//     Drive/Inputs/In/nState1 @bit 4 <-> STM Status/Status/Moving positive
//     Drive/Inputs/In/nState1 @bit 1 <-> STM Status/Status/Ready
//     Drive/Inputs/In/nState1 <-> STM Status/Status/Ready to enable
//     Drive/Inputs/In/nState1 @bit 6 <-> STM Status/Status/Torque reduced
//     Drive/Inputs/In/nState1 @bit 2 <-> STM Status/Status/Warning
//     Drive/Inputs/In/nState2 @bit 3 <-> STM Status/Status/Digital input 1
//     Drive/Inputs/In/nState2 @bit 4 <-> STM Status/Status/Digital input 2
//     Drive/Inputs/In/nState2 @bit 5 <-> STM Status/Status/Sync error
//     Drive/Inputs/In/nState2 @bit 7 <-> STM Status/Status/TxPDO Toggle
//     Drive/Inputs/In/nState4 @bit 1 <-> WcState/InputToggle
//     Drive/Inputs/In/nState4 <-> WcState/WcState
//     Drive/Outputs/Out/nCtrl1 <-> STM Control/Control/Enable
//     Drive/Outputs/Out/nCtrl1 @bit 2 <-> STM Control/Control/Reduce torque
//     Drive/Outputs/Out/nCtrl1 @bit 1 <-> STM Control/Control/Reset
//     Drive/Outputs/Out/nDataOut2[0] <-> STM Velocity/Velocity
//   (this object) <-> PLC Rail (EtherCAT)/Power (EK1200)/PLC Junction 2 (EK1122)/X1 HXR EC1 (EK1100)/EC1 E2 (EK1122)/X1 IM2L0-XTES (EK1100)/IM2L0-EL5042
//     Enc/Inputs/In/nComState @bit 1 <-> WcState/InputToggle
//     Enc/Inputs/In/nComState <-> WcState/WcState
//     Enc/Inputs/In/nDataIn1 <-> FB Inputs Channel 1/Position
//     Enc/Inputs/In/nState1 @bit 12 <-> FB Inputs Channel 1/Status/Diag
//     Enc/Inputs/In/nState1 @bit 1 <-> FB Inputs Channel 1/Status/Error
//     Enc/Inputs/In/nState1 @bit 14 <-> FB Inputs Channel 1/Status/Input cycle counter
//     Enc/Inputs/In/nState1 @bit 2 <-> FB Inputs Channel 1/Status/Ready
//     Enc/Inputs/In/nState1 @bit 13 <-> FB Inputs Channel 1/Status/TxPDO State
//     Enc/Inputs/In/nState1 <-> FB Inputs Channel 1/Status/Warning
//   (this object) <-> PLC Rail (EtherCAT)/Power (EK1200)/PLC Junction 2 (EK1122)/X1 HXR EC1 (EK1100)/EC1 E2 (EK1122)/X1 IM2L0-XTES (EK1100)/IM2L0-EL7041
//     Drive/Inputs/In/nState1 @bit 3 <-> STM Status/Status/Error
//     Drive/Inputs/In/nState1 @bit 5 <-> STM Status/Status/Moving negative
//     Drive/Inputs/In/nState1 @bit 4 <-> STM Status/Status/Moving positive
//     Drive/Inputs/In/nState1 @bit 1 <-> STM Status/Status/Ready
//     Drive/Inputs/In/nState1 <-> STM Status/Status/Ready to enable
//     Drive/Inputs/In/nState1 @bit 6 <-> STM Status/Status/Torque reduced
//     Drive/Inputs/In/nState1 @bit 2 <-> STM Status/Status/Warning
//     Drive/Inputs/In/nState2 @bit 3 <-> STM Status/Status/Digital input 1
//     Drive/Inputs/In/nState2 @bit 4 <-> STM Status/Status/Digital input 2
//     Drive/Inputs/In/nState2 @bit 5 <-> STM Status/Status/Sync error
//     Drive/Inputs/In/nState2 @bit 7 <-> STM Status/Status/TxPDO Toggle
//     Drive/Inputs/In/nState4 @bit 1 <-> WcState/InputToggle
//     Drive/Inputs/In/nState4 <-> WcState/WcState
//     Drive/Outputs/Out/nCtrl1 <-> STM Control/Control/Enable
//     Drive/Outputs/Out/nCtrl1 @bit 2 <-> STM Control/Control/Reduce torque
//     Drive/Outputs/Out/nCtrl1 @bit 1 <-> STM Control/Control/Reset
//     Drive/Outputs/Out/nDataOut2[0] <-> STM Velocity/Velocity
//   (this object) <-> PLC Rail (EtherCAT)/Power (EK1200)/PLC Junction 2 (EK1122)/X1 HXR EC1 (EK1100)/EC1 E2 (EK1122)/X1 IM2L0-XTES (EK1100)/IM2L0-EL7342
//     Drive/Inputs/In/nState1 @bit 3 <-> DCM Status Channel 1/Status/Error
//     Drive/Inputs/In/nState1 @bit 3 <-> DCM Status Channel 2/Status/Error
//     Drive/Inputs/In/nState1 @bit 5 <-> DCM Status Channel 1/Status/Moving negative
//     Drive/Inputs/In/nState1 @bit 5 <-> DCM Status Channel 2/Status/Moving negative
//     Drive/Inputs/In/nState1 @bit 4 <-> DCM Status Channel 1/Status/Moving positive
//     Drive/Inputs/In/nState1 @bit 4 <-> DCM Status Channel 2/Status/Moving positive
//     Drive/Inputs/In/nState1 @bit 1 <-> DCM Status Channel 1/Status/Ready
//     Drive/Inputs/In/nState1 @bit 1 <-> DCM Status Channel 2/Status/Ready
//     Drive/Inputs/In/nState1 <-> DCM Status Channel 1/Status/Ready to enable
//     Drive/Inputs/In/nState1 <-> DCM Status Channel 2/Status/Ready to enable
//     Drive/Inputs/In/nState1 @bit 6 <-> DCM Status Channel 1/Status/Torque reduced
//     Drive/Inputs/In/nState1 @bit 6 <-> DCM Status Channel 2/Status/Torque reduced
//     Drive/Inputs/In/nState1 @bit 2 <-> DCM Status Channel 1/Status/Warning
//     Drive/Inputs/In/nState1 @bit 2 <-> DCM Status Channel 2/Status/Warning
//     Drive/Inputs/In/nState2 @bit 3 <-> DCM Status Channel 1/Status/Digital input 1
//     Drive/Inputs/In/nState2 @bit 4 <-> DCM Status Channel 1/Status/Digital input 2
//     Drive/Inputs/In/nState2 @bit 3 <-> DCM Status Channel 2/Status/Digital input 1
//     Drive/Inputs/In/nState2 @bit 4 <-> DCM Status Channel 2/Status/Digital input 2
//     Drive/Inputs/In/nState2 @bit 5 <-> DCM Status Channel 1/Status/Sync error
//     Drive/Inputs/In/nState2 @bit 5 <-> DCM Status Channel 2/Status/Sync error
//     Drive/Inputs/In/nState2 @bit 7 <-> DCM Status Channel 1/Status/TxPDO Toggle
//     Drive/Inputs/In/nState2 @bit 7 <-> DCM Status Channel 2/Status/TxPDO Toggle
//     Drive/Inputs/In/nState4 @bit 1 <-> WcState/InputToggle
//     Drive/Inputs/In/nState4 <-> WcState/WcState
//     Drive/Outputs/Out/nCtrl1 <-> DCM Control Channel 1/Control/Enable
//     Drive/Outputs/Out/nCtrl1 <-> DCM Control Channel 2/Control/Enable
//     Drive/Outputs/Out/nCtrl1 @bit 2 <-> DCM Control Channel 1/Control/Reduce torque
//     Drive/Outputs/Out/nCtrl1 @bit 2 <-> DCM Control Channel 2/Control/Reduce torque
//     Drive/Outputs/Out/nCtrl1 @bit 1 <-> DCM Control Channel 1/Control/Reset
//     Drive/Outputs/Out/nCtrl1 @bit 1 <-> DCM Control Channel 2/Control/Reset
//     Drive/Outputs/Out/nCtrl1 @bit 3 <-> DCM Control Channel 1/Control/Threshold active
//     Drive/Outputs/Out/nCtrl1 @bit 3 <-> DCM Control Channel 2/Control/Threshold active
//     Drive/Outputs/Out/nDataOut2[0] <-> DCM Velocity Channel 1/Velocity
//     Drive/Outputs/Out/nDataOut2[0] <-> DCM Velocity Channel 2/Velocity
//     Enc/Inputs/In/nDataIn1[0] <-> ENC Status compact Channel 1/Counter value
//     Enc/Inputs/In/nDataIn1[0] <-> ENC Status compact Channel 2/Counter value
//     Enc/Inputs/In/nDataIn2[0] <-> ENC Status compact Channel 1/Latch value
//     Enc/Inputs/In/nDataIn2[0] <-> ENC Status compact Channel 2/Latch value
//     Enc/Inputs/In/nState1 @bit 4 <-> ENC Status compact Channel 1/Status/Counter overflow
//     Enc/Inputs/In/nState1 @bit 4 <-> ENC Status compact Channel 2/Status/Counter overflow
//     Enc/Inputs/In/nState1 @bit 3 <-> ENC Status compact Channel 1/Status/Counter underflow
//     Enc/Inputs/In/nState1 @bit 3 <-> ENC Status compact Channel 2/Status/Counter underflow
//     Enc/Inputs/In/nState1 @bit 7 <-> ENC Status compact Channel 1/Status/Extrapolation stall
//     Enc/Inputs/In/nState1 @bit 7 <-> ENC Status compact Channel 2/Status/Extrapolation stall
//     Enc/Inputs/In/nState1 @bit 1 <-> ENC Status compact Channel 1/Status/Latch extern valid
//     Enc/Inputs/In/nState1 @bit 1 <-> ENC Status compact Channel 2/Status/Latch extern valid
//     Enc/Inputs/In/nState1 @bit 2 <-> ENC Status compact Channel 1/Status/Set counter done
//     Enc/Inputs/In/nState1 @bit 2 <-> ENC Status compact Channel 2/Status/Set counter done
//     Enc/Inputs/In/nState2 @bit 4 <-> ENC Status compact Channel 1/Status/Status of extern latch
//     Enc/Inputs/In/nState2 @bit 4 <-> ENC Status compact Channel 2/Status/Status of extern latch
//     Enc/Inputs/In/nState2 <-> ENC Status compact Channel 1/Status/Status of input A
//     Enc/Inputs/In/nState2 <-> ENC Status compact Channel 2/Status/Status of input A
//     Enc/Inputs/In/nState2 @bit 1 <-> ENC Status compact Channel 1/Status/Status of input B
//     Enc/Inputs/In/nState2 @bit 1 <-> ENC Status compact Channel 2/Status/Status of input B
//     Enc/Inputs/In/nState2 @bit 5 <-> ENC Status compact Channel 1/Status/Sync error
//     Enc/Inputs/In/nState2 @bit 5 <-> ENC Status compact Channel 2/Status/Sync error
//     Enc/Inputs/In/nState2 @bit 7 <-> ENC Status compact Channel 1/Status/TxPDO Toggle
//     Enc/Inputs/In/nState2 @bit 7 <-> ENC Status compact Channel 2/Status/TxPDO Toggle
//     Enc/Inputs/In/nState4 @bit 1 <-> WcState/InputToggle
//     Enc/Inputs/In/nState4 <-> WcState/WcState
//     Enc/Outputs/Out/nCtrl1 @bit 3 <-> ENC Control compact Channel 1/Control/Enable latch extern on negative edge
//     Enc/Outputs/Out/nCtrl1 @bit 3 <-> ENC Control compact Channel 2/Control/Enable latch extern on negative edge
//     Enc/Outputs/Out/nCtrl1 @bit 1 <-> ENC Control compact Channel 1/Control/Enable latch extern on positive edge
//     Enc/Outputs/Out/nCtrl1 @bit 1 <-> ENC Control compact Channel 2/Control/Enable latch extern on positive edge
//     Enc/Outputs/Out/nCtrl1 @bit 2 <-> ENC Control compact Channel 1/Control/Set counter
//     Enc/Outputs/Out/nCtrl1 @bit 2 <-> ENC Control compact Channel 2/Control/Set counter
//     Enc/Outputs/Out/nDataOut1[0] <-> ENC Control compact Channel 1/Set counter value
//     Enc/Outputs/Out/nDataOut1[0] <-> ENC Control compact Channel 2/Set counter value
//   (this object) <-> PLC Rail (EtherCAT)/Power (EK1200)/PLC Junction 2 (EK1122)/X2 HXR EC2 (EK1100)/EC2 E1 (EK1122)/X1 IM3L0-PPM (EK1100)/IM3L0-EL5042
//     Enc/Inputs/In/nComState @bit 1 <-> WcState/InputToggle
//     Enc/Inputs/In/nComState <-> WcState/WcState
//     Enc/Inputs/In/nDataIn1 <-> FB Inputs Channel 1/Position
//     Enc/Inputs/In/nState1 @bit 12 <-> FB Inputs Channel 1/Status/Diag
//     Enc/Inputs/In/nState1 @bit 1 <-> FB Inputs Channel 1/Status/Error
//     Enc/Inputs/In/nState1 @bit 14 <-> FB Inputs Channel 1/Status/Input cycle counter
//     Enc/Inputs/In/nState1 @bit 2 <-> FB Inputs Channel 1/Status/Ready
//     Enc/Inputs/In/nState1 @bit 13 <-> FB Inputs Channel 1/Status/TxPDO State
//     Enc/Inputs/In/nState1 <-> FB Inputs Channel 1/Status/Warning
//   (this object) <-> PLC Rail (EtherCAT)/Power (EK1200)/PLC Junction 2 (EK1122)/X2 HXR EC2 (EK1100)/EC2 E1 (EK1122)/X1 IM3L0-PPM (EK1100)/IM3L0-EL7041
//     Drive/Inputs/In/nState1 @bit 3 <-> STM Status/Status/Error
//     Drive/Inputs/In/nState1 @bit 5 <-> STM Status/Status/Moving negative
//     Drive/Inputs/In/nState1 @bit 4 <-> STM Status/Status/Moving positive
//     Drive/Inputs/In/nState1 @bit 1 <-> STM Status/Status/Ready
//     Drive/Inputs/In/nState1 <-> STM Status/Status/Ready to enable
//     Drive/Inputs/In/nState1 @bit 6 <-> STM Status/Status/Torque reduced
//     Drive/Inputs/In/nState1 @bit 2 <-> STM Status/Status/Warning
//     Drive/Inputs/In/nState2 @bit 3 <-> STM Status/Status/Digital input 1
//     Drive/Inputs/In/nState2 @bit 4 <-> STM Status/Status/Digital input 2
//     Drive/Inputs/In/nState2 @bit 5 <-> STM Status/Status/Sync error
//     Drive/Inputs/In/nState2 @bit 7 <-> STM Status/Status/TxPDO Toggle
//     Drive/Inputs/In/nState4 @bit 1 <-> WcState/InputToggle
//     Drive/Inputs/In/nState4 <-> WcState/WcState
//     Drive/Outputs/Out/nCtrl1 <-> STM Control/Control/Enable
//     Drive/Outputs/Out/nCtrl1 @bit 2 <-> STM Control/Control/Reduce torque
//     Drive/Outputs/Out/nCtrl1 @bit 1 <-> STM Control/Control/Reset
//     Drive/Outputs/Out/nDataOut2[0] <-> STM Velocity/Velocity
//   (this object) <-> PLC Rail (EtherCAT)/Power (EK1200)/PLC Junction 2 (EK1122)/X2 HXR EC2 (EK1100)/EC2 E2 (EK1122)/X1 IM4L0-XTES (EK1100)/IM4L0-EL5042
//     Enc/Inputs/In/nComState @bit 1 <-> WcState/InputToggle
//     Enc/Inputs/In/nComState <-> WcState/WcState
//     Enc/Inputs/In/nDataIn1 <-> FB Inputs Channel 1/Position
//     Enc/Inputs/In/nState1 @bit 12 <-> FB Inputs Channel 1/Status/Diag
//     Enc/Inputs/In/nState1 @bit 1 <-> FB Inputs Channel 1/Status/Error
//     Enc/Inputs/In/nState1 @bit 14 <-> FB Inputs Channel 1/Status/Input cycle counter
//     Enc/Inputs/In/nState1 @bit 2 <-> FB Inputs Channel 1/Status/Ready
//     Enc/Inputs/In/nState1 @bit 13 <-> FB Inputs Channel 1/Status/TxPDO State
//     Enc/Inputs/In/nState1 <-> FB Inputs Channel 1/Status/Warning
//   (this object) <-> PLC Rail (EtherCAT)/Power (EK1200)/PLC Junction 2 (EK1122)/X2 HXR EC2 (EK1100)/EC2 E2 (EK1122)/X1 IM4L0-XTES (EK1100)/IM4L0-EL7041
//     Drive/Inputs/In/nState1 @bit 3 <-> STM Status/Status/Error
//     Drive/Inputs/In/nState1 @bit 5 <-> STM Status/Status/Moving negative
//     Drive/Inputs/In/nState1 @bit 4 <-> STM Status/Status/Moving positive
//     Drive/Inputs/In/nState1 @bit 1 <-> STM Status/Status/Ready
//     Drive/Inputs/In/nState1 <-> STM Status/Status/Ready to enable
//     Drive/Inputs/In/nState1 @bit 6 <-> STM Status/Status/Torque reduced
//     Drive/Inputs/In/nState1 @bit 2 <-> STM Status/Status/Warning
//     Drive/Inputs/In/nState2 @bit 3 <-> STM Status/Status/Digital input 1
//     Drive/Inputs/In/nState2 @bit 4 <-> STM Status/Status/Digital input 2
//     Drive/Inputs/In/nState2 @bit 5 <-> STM Status/Status/Sync error
//     Drive/Inputs/In/nState2 @bit 7 <-> STM Status/Status/TxPDO Toggle
//     Drive/Inputs/In/nState4 @bit 1 <-> WcState/InputToggle
//     Drive/Inputs/In/nState4 <-> WcState/WcState
//     Drive/Outputs/Out/nCtrl1 <-> STM Control/Control/Enable
//     Drive/Outputs/Out/nCtrl1 @bit 2 <-> STM Control/Control/Reduce torque
//     Drive/Outputs/Out/nCtrl1 @bit 1 <-> STM Control/Control/Reset
//     Drive/Outputs/Out/nDataOut2[0] <-> STM Velocity/Velocity
//   (this object) <-> PLC Rail (EtherCAT)/Power (EK1200)/PLC Junction 2 (EK1122)/X2 HXR EC2 (EK1100)/EC2 E2 (EK1122)/X1 IM4L0-XTES (EK1100)/IM4L0-EL7342
//     Drive/Inputs/In/nState1 @bit 3 <-> DCM Status Channel 1/Status/Error
//     Drive/Inputs/In/nState1 @bit 3 <-> DCM Status Channel 2/Status/Error
//     Drive/Inputs/In/nState1 @bit 5 <-> DCM Status Channel 1/Status/Moving negative
//     Drive/Inputs/In/nState1 @bit 5 <-> DCM Status Channel 2/Status/Moving negative
//     Drive/Inputs/In/nState1 @bit 4 <-> DCM Status Channel 1/Status/Moving positive
//     Drive/Inputs/In/nState1 @bit 4 <-> DCM Status Channel 2/Status/Moving positive
//     Drive/Inputs/In/nState1 @bit 1 <-> DCM Status Channel 1/Status/Ready
//     Drive/Inputs/In/nState1 @bit 1 <-> DCM Status Channel 2/Status/Ready
//     Drive/Inputs/In/nState1 <-> DCM Status Channel 1/Status/Ready to enable
//     Drive/Inputs/In/nState1 <-> DCM Status Channel 2/Status/Ready to enable
//     Drive/Inputs/In/nState1 @bit 6 <-> DCM Status Channel 1/Status/Torque reduced
//     Drive/Inputs/In/nState1 @bit 6 <-> DCM Status Channel 2/Status/Torque reduced
//     Drive/Inputs/In/nState1 @bit 2 <-> DCM Status Channel 1/Status/Warning
//     Drive/Inputs/In/nState1 @bit 2 <-> DCM Status Channel 2/Status/Warning
//     Drive/Inputs/In/nState2 @bit 3 <-> DCM Status Channel 1/Status/Digital input 1
//     Drive/Inputs/In/nState2 @bit 4 <-> DCM Status Channel 1/Status/Digital input 2
//     Drive/Inputs/In/nState2 @bit 3 <-> DCM Status Channel 2/Status/Digital input 1
//     Drive/Inputs/In/nState2 @bit 4 <-> DCM Status Channel 2/Status/Digital input 2
//     Drive/Inputs/In/nState2 @bit 5 <-> DCM Status Channel 1/Status/Sync error
//     Drive/Inputs/In/nState2 @bit 5 <-> DCM Status Channel 2/Status/Sync error
//     Drive/Inputs/In/nState2 @bit 7 <-> DCM Status Channel 1/Status/TxPDO Toggle
//     Drive/Inputs/In/nState2 @bit 7 <-> DCM Status Channel 2/Status/TxPDO Toggle
//     Drive/Inputs/In/nState4 @bit 1 <-> WcState/InputToggle
//     Drive/Inputs/In/nState4 <-> WcState/WcState
//     Drive/Outputs/Out/nCtrl1 <-> DCM Control Channel 1/Control/Enable
//     Drive/Outputs/Out/nCtrl1 <-> DCM Control Channel 2/Control/Enable
//     Drive/Outputs/Out/nCtrl1 @bit 2 <-> DCM Control Channel 1/Control/Reduce torque
//     Drive/Outputs/Out/nCtrl1 @bit 2 <-> DCM Control Channel 2/Control/Reduce torque
//     Drive/Outputs/Out/nCtrl1 @bit 1 <-> DCM Control Channel 1/Control/Reset
//     Drive/Outputs/Out/nCtrl1 @bit 1 <-> DCM Control Channel 2/Control/Reset
//     Drive/Outputs/Out/nCtrl1 @bit 3 <-> DCM Control Channel 1/Control/Threshold active
//     Drive/Outputs/Out/nCtrl1 @bit 3 <-> DCM Control Channel 2/Control/Threshold active
//     Drive/Outputs/Out/nDataOut2[0] <-> DCM Velocity Channel 1/Velocity
//     Drive/Outputs/Out/nDataOut2[0] <-> DCM Velocity Channel 2/Velocity
//     Enc/Inputs/In/nDataIn1[0] <-> ENC Status compact Channel 1/Counter value
//     Enc/Inputs/In/nDataIn1[0] <-> ENC Status compact Channel 2/Counter value
//     Enc/Inputs/In/nDataIn2[0] <-> ENC Status compact Channel 1/Latch value
//     Enc/Inputs/In/nDataIn2[0] <-> ENC Status compact Channel 2/Latch value
//     Enc/Inputs/In/nState1 @bit 4 <-> ENC Status compact Channel 1/Status/Counter overflow
//     Enc/Inputs/In/nState1 @bit 4 <-> ENC Status compact Channel 2/Status/Counter overflow
//     Enc/Inputs/In/nState1 @bit 3 <-> ENC Status compact Channel 1/Status/Counter underflow
//     Enc/Inputs/In/nState1 @bit 3 <-> ENC Status compact Channel 2/Status/Counter underflow
//     Enc/Inputs/In/nState1 @bit 7 <-> ENC Status compact Channel 1/Status/Extrapolation stall
//     Enc/Inputs/In/nState1 @bit 7 <-> ENC Status compact Channel 2/Status/Extrapolation stall
//     Enc/Inputs/In/nState1 @bit 1 <-> ENC Status compact Channel 1/Status/Latch extern valid
//     Enc/Inputs/In/nState1 @bit 1 <-> ENC Status compact Channel 2/Status/Latch extern valid
//     Enc/Inputs/In/nState1 @bit 2 <-> ENC Status compact Channel 1/Status/Set counter done
//     Enc/Inputs/In/nState1 @bit 2 <-> ENC Status compact Channel 2/Status/Set counter done
//     Enc/Inputs/In/nState2 @bit 4 <-> ENC Status compact Channel 1/Status/Status of extern latch
//     Enc/Inputs/In/nState2 @bit 4 <-> ENC Status compact Channel 2/Status/Status of extern latch
//     Enc/Inputs/In/nState2 <-> ENC Status compact Channel 1/Status/Status of input A
//     Enc/Inputs/In/nState2 <-> ENC Status compact Channel 2/Status/Status of input A
//     Enc/Inputs/In/nState2 @bit 1 <-> ENC Status compact Channel 1/Status/Status of input B
//     Enc/Inputs/In/nState2 @bit 1 <-> ENC Status compact Channel 2/Status/Status of input B
//     Enc/Inputs/In/nState2 @bit 5 <-> ENC Status compact Channel 1/Status/Sync error
//     Enc/Inputs/In/nState2 @bit 5 <-> ENC Status compact Channel 2/Status/Sync error
//     Enc/Inputs/In/nState2 @bit 7 <-> ENC Status compact Channel 1/Status/TxPDO Toggle
//     Enc/Inputs/In/nState2 @bit 7 <-> ENC Status compact Channel 2/Status/TxPDO Toggle
//     Enc/Inputs/In/nState4 @bit 1 <-> WcState/InputToggle
//     Enc/Inputs/In/nState4 <-> WcState/WcState
//     Enc/Outputs/Out/nCtrl1 @bit 3 <-> ENC Control compact Channel 1/Control/Enable latch extern on negative edge
//     Enc/Outputs/Out/nCtrl1 @bit 3 <-> ENC Control compact Channel 2/Control/Enable latch extern on negative edge
//     Enc/Outputs/Out/nCtrl1 @bit 1 <-> ENC Control compact Channel 1/Control/Enable latch extern on positive edge
//     Enc/Outputs/Out/nCtrl1 @bit 1 <-> ENC Control compact Channel 2/Control/Enable latch extern on positive edge
//     Enc/Outputs/Out/nCtrl1 @bit 2 <-> ENC Control compact Channel 1/Control/Set counter
//     Enc/Outputs/Out/nCtrl1 @bit 2 <-> ENC Control compact Channel 2/Control/Set counter
//     Enc/Outputs/Out/nDataOut1[0] <-> ENC Control compact Channel 1/Set counter value
//     Enc/Outputs/Out/nDataOut1[0] <-> ENC Control compact Channel 2/Set counter value
//   (this object) <-> PLC Rail (EtherCAT)/Power (EK1200)/PLC Junction 2 (EK1122)/X1 HXR EC1 (EK1100)/EC1 E3 (EK1122)/X1 PF1L0-WFS (EK1100)/PF1L0-EL5042
//     Enc/Inputs/In/nComState @bit 1 <-> WcState/InputToggle
//     Enc/Inputs/In/nComState <-> WcState/WcState
//     Enc/Inputs/In/nDataIn1 <-> FB Inputs Channel 2/Position
//     Enc/Inputs/In/nDataIn1 <-> FB Inputs Channel 1/Position
//     Enc/Inputs/In/nState1 @bit 12 <-> FB Inputs Channel 2/Status/Diag
//     Enc/Inputs/In/nState1 @bit 12 <-> FB Inputs Channel 1/Status/Diag
//     Enc/Inputs/In/nState1 @bit 1 <-> FB Inputs Channel 2/Status/Error
//     Enc/Inputs/In/nState1 @bit 1 <-> FB Inputs Channel 1/Status/Error
//     Enc/Inputs/In/nState1 @bit 14 <-> FB Inputs Channel 2/Status/Input cycle counter
//     Enc/Inputs/In/nState1 @bit 14 <-> FB Inputs Channel 1/Status/Input cycle counter
//     Enc/Inputs/In/nState1 @bit 2 <-> FB Inputs Channel 2/Status/Ready
//     Enc/Inputs/In/nState1 @bit 2 <-> FB Inputs Channel 1/Status/Ready
//     Enc/Inputs/In/nState1 @bit 13 <-> FB Inputs Channel 2/Status/TxPDO State
//     Enc/Inputs/In/nState1 @bit 13 <-> FB Inputs Channel 1/Status/TxPDO State
//     Enc/Inputs/In/nState1 <-> FB Inputs Channel 2/Status/Warning
//     Enc/Inputs/In/nState1 <-> FB Inputs Channel 1/Status/Warning
//   (this object) <-> PLC Rail (EtherCAT)/Power (EK1200)/PLC Junction 2 (EK1122)/X1 HXR EC1 (EK1100)/EC1 E3 (EK1122)/X1 PF1L0-WFS (EK1100)/PF1L0-EL7041-01
//     Drive/Inputs/In/nState1 @bit 3 <-> STM Status/Status/Error
//     Drive/Inputs/In/nState1 @bit 5 <-> STM Status/Status/Moving negative
//     Drive/Inputs/In/nState1 @bit 4 <-> STM Status/Status/Moving positive
//     Drive/Inputs/In/nState1 @bit 1 <-> STM Status/Status/Ready
//     Drive/Inputs/In/nState1 <-> STM Status/Status/Ready to enable
//     Drive/Inputs/In/nState1 @bit 6 <-> STM Status/Status/Torque reduced
//     Drive/Inputs/In/nState1 @bit 2 <-> STM Status/Status/Warning
//     Drive/Inputs/In/nState2 @bit 3 <-> STM Status/Status/Digital input 1
//     Drive/Inputs/In/nState2 @bit 4 <-> STM Status/Status/Digital input 2
//     Drive/Inputs/In/nState2 @bit 5 <-> STM Status/Status/Sync error
//     Drive/Inputs/In/nState2 @bit 7 <-> STM Status/Status/TxPDO Toggle
//     Drive/Inputs/In/nState4 @bit 1 <-> WcState/InputToggle
//     Drive/Inputs/In/nState4 <-> WcState/WcState
//     Drive/Outputs/Out/nCtrl1 <-> STM Control/Control/Enable
//     Drive/Outputs/Out/nCtrl1 @bit 2 <-> STM Control/Control/Reduce torque
//     Drive/Outputs/Out/nCtrl1 @bit 1 <-> STM Control/Control/Reset
//     Drive/Outputs/Out/nDataOut2[0] <-> STM Velocity/Velocity
//   (this object) <-> PLC Rail (EtherCAT)/Power (EK1200)/PLC Junction 2 (EK1122)/X1 HXR EC1 (EK1100)/EC1 E3 (EK1122)/X1 PF1L0-WFS (EK1100)/PF1L0-EL7041-02
//     Drive/Inputs/In/nState1 @bit 3 <-> STM Status/Status/Error
//     Drive/Inputs/In/nState1 @bit 5 <-> STM Status/Status/Moving negative
//     Drive/Inputs/In/nState1 @bit 4 <-> STM Status/Status/Moving positive
//     Drive/Inputs/In/nState1 @bit 1 <-> STM Status/Status/Ready
//     Drive/Inputs/In/nState1 <-> STM Status/Status/Ready to enable
//     Drive/Inputs/In/nState1 @bit 6 <-> STM Status/Status/Torque reduced
//     Drive/Inputs/In/nState1 @bit 2 <-> STM Status/Status/Warning
//     Drive/Inputs/In/nState2 @bit 3 <-> STM Status/Status/Digital input 1
//     Drive/Inputs/In/nState2 @bit 4 <-> STM Status/Status/Digital input 2
//     Drive/Inputs/In/nState2 @bit 5 <-> STM Status/Status/Sync error
//     Drive/Inputs/In/nState2 @bit 7 <-> STM Status/Status/TxPDO Toggle
//     Drive/Inputs/In/nState4 @bit 1 <-> WcState/InputToggle
//     Drive/Inputs/In/nState4 <-> WcState/WcState
//     Drive/Outputs/Out/nCtrl1 <-> STM Control/Control/Enable
//     Drive/Outputs/Out/nCtrl1 @bit 2 <-> STM Control/Control/Reduce torque
//     Drive/Outputs/Out/nCtrl1 @bit 1 <-> STM Control/Control/Reset
//     Drive/Outputs/Out/nDataOut2[0] <-> STM Velocity/Velocity
//   (this object) <-> PLC Rail (EtherCAT)/Power (EK1200)/PLC Junction 1 (EK1122)/X1 RTDSL0 (EK1100)/RTDSL0-EL7041-01
//     Drive/Inputs/In/nState1 @bit 3 <-> STM Status/Status/Error
//     Drive/Inputs/In/nState1 @bit 5 <-> STM Status/Status/Moving negative
//     Drive/Inputs/In/nState1 @bit 4 <-> STM Status/Status/Moving positive
//     Drive/Inputs/In/nState1 @bit 1 <-> STM Status/Status/Ready
//     Drive/Inputs/In/nState1 <-> STM Status/Status/Ready to enable
//     Drive/Inputs/In/nState1 @bit 6 <-> STM Status/Status/Torque reduced
//     Drive/Inputs/In/nState1 @bit 2 <-> STM Status/Status/Warning
//     Drive/Inputs/In/nState2 @bit 3 <-> STM Status/Status/Digital input 1
//     Drive/Inputs/In/nState2 @bit 4 <-> STM Status/Status/Digital input 2
//     Drive/Inputs/In/nState2 @bit 5 <-> STM Status/Status/Sync error
//     Drive/Inputs/In/nState2 @bit 7 <-> STM Status/Status/TxPDO Toggle
//     Drive/Inputs/In/nState4 @bit 1 <-> WcState/InputToggle
//     Drive/Inputs/In/nState4 <-> WcState/WcState
//     Drive/Outputs/Out/nCtrl1 <-> STM Control/Control/Enable
//     Drive/Outputs/Out/nCtrl1 @bit 2 <-> STM Control/Control/Reduce torque
//     Drive/Outputs/Out/nCtrl1 @bit 1 <-> STM Control/Control/Reset
//     Drive/Outputs/Out/nDataOut2[0] <-> STM Velocity/Velocity
//     Enc/Inputs/In/nDataIn1[0] <-> ENC Status compact/Counter value
//     Enc/Inputs/In/nDataIn2[0] <-> ENC Status compact/Latch value
//     Enc/Inputs/In/nState1 @bit 4 <-> ENC Status compact/Status/Counter overflow
//     Enc/Inputs/In/nState1 @bit 3 <-> ENC Status compact/Status/Counter underflow
//     Enc/Inputs/In/nState1 @bit 7 <-> ENC Status compact/Status/Extrapolation stall
//     Enc/Inputs/In/nState1 <-> ENC Status compact/Status/Latch C valid
//     Enc/Inputs/In/nState1 @bit 1 <-> ENC Status compact/Status/Latch extern valid
//     Enc/Inputs/In/nState1 @bit 2 <-> ENC Status compact/Status/Set counter done
//     Enc/Inputs/In/nState2 @bit 4 <-> ENC Status compact/Status/Status of extern latch
//     Enc/Inputs/In/nState2 <-> ENC Status compact/Status/Status of input A
//     Enc/Inputs/In/nState2 @bit 1 <-> ENC Status compact/Status/Status of input B
//     Enc/Inputs/In/nState2 @bit 2 <-> ENC Status compact/Status/Status of input C
//     Enc/Inputs/In/nState2 @bit 5 <-> ENC Status compact/Status/Sync error
//     Enc/Inputs/In/nState2 @bit 7 <-> ENC Status compact/Status/TxPDO Toggle
//     Enc/Inputs/In/nState4 @bit 1 <-> WcState/InputToggle
//     Enc/Inputs/In/nState4 <-> WcState/WcState
//     Enc/Outputs/Out/nCtrl1 <-> ENC Control compact/Control/Enable latch C
//     Enc/Outputs/Out/nCtrl1 @bit 3 <-> ENC Control compact/Control/Enable latch extern on negative edge
//     Enc/Outputs/Out/nCtrl1 @bit 1 <-> ENC Control compact/Control/Enable latch extern on positive edge
//     Enc/Outputs/Out/nCtrl1 @bit 2 <-> ENC Control compact/Control/Set counter
//     Enc/Outputs/Out/nDataOut1[0] <-> ENC Control compact/Set counter value
//   (this object) <-> PLC Rail (EtherCAT)/Power (EK1200)/PLC Junction 1 (EK1122)/X1 RTDSL0 (EK1100)/RTDSL0-EL7041-05
//     Drive/Inputs/In/nState1 @bit 3 <-> STM Status/Status/Error
//     Drive/Inputs/In/nState1 @bit 5 <-> STM Status/Status/Moving negative
//     Drive/Inputs/In/nState1 @bit 4 <-> STM Status/Status/Moving positive
//     Drive/Inputs/In/nState1 @bit 1 <-> STM Status/Status/Ready
//     Drive/Inputs/In/nState1 <-> STM Status/Status/Ready to enable
//     Drive/Inputs/In/nState1 @bit 6 <-> STM Status/Status/Torque reduced
//     Drive/Inputs/In/nState1 @bit 2 <-> STM Status/Status/Warning
//     Drive/Inputs/In/nState2 @bit 3 <-> STM Status/Status/Digital input 1
//     Drive/Inputs/In/nState2 @bit 4 <-> STM Status/Status/Digital input 2
//     Drive/Inputs/In/nState2 @bit 5 <-> STM Status/Status/Sync error
//     Drive/Inputs/In/nState2 @bit 7 <-> STM Status/Status/TxPDO Toggle
//     Drive/Inputs/In/nState4 @bit 1 <-> WcState/InputToggle
//     Drive/Inputs/In/nState4 <-> WcState/WcState
//     Drive/Outputs/Out/nCtrl1 <-> STM Control/Control/Enable
//     Drive/Outputs/Out/nCtrl1 @bit 2 <-> STM Control/Control/Reduce torque
//     Drive/Outputs/Out/nCtrl1 @bit 1 <-> STM Control/Control/Reset
//     Drive/Outputs/Out/nDataOut2[0] <-> STM Velocity/Velocity
//   (this object) <-> PLC Rail (EtherCAT)/Power (EK1200)/PLC Junction 1 (EK1122)/X1 RTDSL0 (EK1100)/Term 113 (EL3054)
//     Enc/Inputs/In/nDataIn1[0] <-> AI Standard Channel 1/Value
//     Enc/Inputs/In/nState4 @bit 1 <-> WcState/InputToggle
//     Enc/Inputs/In/nState4 <-> WcState/WcState
//   (this object) <-> PLC Rail (EtherCAT)/Power (EK1200)/PLC Junction 2 (EK1122)/X1 HXR EC1 (EK1100)/EC1 E1 (EK1122)/X1 SL1L0-Power (EK1100)/SL1L0-EL5042-E2
//     Enc/Inputs/In/nComState @bit 1 <-> WcState/InputToggle
//     Enc/Inputs/In/nComState <-> WcState/WcState
//     Enc/Inputs/In/nDataIn1 <-> FB Inputs Channel 1/Position
//     Enc/Inputs/In/nDataIn1 <-> FB Inputs Channel 2/Position
//     Enc/Inputs/In/nState1 @bit 12 <-> FB Inputs Channel 1/Status/Diag
//     Enc/Inputs/In/nState1 @bit 12 <-> FB Inputs Channel 2/Status/Diag
//     Enc/Inputs/In/nState1 @bit 1 <-> FB Inputs Channel 1/Status/Error
//     Enc/Inputs/In/nState1 @bit 1 <-> FB Inputs Channel 2/Status/Error
//     Enc/Inputs/In/nState1 @bit 14 <-> FB Inputs Channel 1/Status/Input cycle counter
//     Enc/Inputs/In/nState1 @bit 14 <-> FB Inputs Channel 2/Status/Input cycle counter
//     Enc/Inputs/In/nState1 @bit 2 <-> FB Inputs Channel 1/Status/Ready
//     Enc/Inputs/In/nState1 @bit 2 <-> FB Inputs Channel 2/Status/Ready
//     Enc/Inputs/In/nState1 @bit 13 <-> FB Inputs Channel 1/Status/TxPDO State
//     Enc/Inputs/In/nState1 @bit 13 <-> FB Inputs Channel 2/Status/TxPDO State
//     Enc/Inputs/In/nState1 <-> FB Inputs Channel 1/Status/Warning
//     Enc/Inputs/In/nState1 <-> FB Inputs Channel 2/Status/Warning
//   (this object) <-> PLC Rail (EtherCAT)/Power (EK1200)/PLC Junction 2 (EK1122)/X1 HXR EC1 (EK1100)/EC1 E1 (EK1122)/X1 SL1L0-Power (EK1100)/SL1L0-EL7041-E1
//     Drive/Inputs/In/nState1 @bit 3 <-> STM Status/Status/Error
//     Drive/Inputs/In/nState1 @bit 5 <-> STM Status/Status/Moving negative
//     Drive/Inputs/In/nState1 @bit 4 <-> STM Status/Status/Moving positive
//     Drive/Inputs/In/nState1 @bit 1 <-> STM Status/Status/Ready
//     Drive/Inputs/In/nState1 <-> STM Status/Status/Ready to enable
//     Drive/Inputs/In/nState1 @bit 6 <-> STM Status/Status/Torque reduced
//     Drive/Inputs/In/nState1 @bit 2 <-> STM Status/Status/Warning
//     Drive/Inputs/In/nState2 @bit 3 <-> STM Status/Status/Digital input 1
//     Drive/Inputs/In/nState2 @bit 4 <-> STM Status/Status/Digital input 2
//     Drive/Inputs/In/nState2 @bit 5 <-> STM Status/Status/Sync error
//     Drive/Inputs/In/nState2 @bit 7 <-> STM Status/Status/TxPDO Toggle
//     Drive/Inputs/In/nState4 @bit 1 <-> WcState/InputToggle
//     Drive/Inputs/In/nState4 <-> WcState/WcState
//     Drive/Outputs/Out/nCtrl1 <-> STM Control/Control/Enable
//     Drive/Outputs/Out/nCtrl1 @bit 2 <-> STM Control/Control/Reduce torque
//     Drive/Outputs/Out/nCtrl1 @bit 1 <-> STM Control/Control/Reset
//     Drive/Outputs/Out/nDataOut2[0] <-> STM Velocity/Velocity
//   (this object) <-> PLC Rail (EtherCAT)/Power (EK1200)/PLC Junction 2 (EK1122)/X1 HXR EC1 (EK1100)/EC1 E1 (EK1122)/X1 SL1L0-Power (EK1100)/SL1L0-EL7041-E3
//     Drive/Inputs/In/nState1 @bit 3 <-> STM Status/Status/Error
//     Drive/Inputs/In/nState1 @bit 5 <-> STM Status/Status/Moving negative
//     Drive/Inputs/In/nState1 @bit 4 <-> STM Status/Status/Moving positive
//     Drive/Inputs/In/nState1 @bit 1 <-> STM Status/Status/Ready
//     Drive/Inputs/In/nState1 <-> STM Status/Status/Ready to enable
//     Drive/Inputs/In/nState1 @bit 6 <-> STM Status/Status/Torque reduced
//     Drive/Inputs/In/nState1 @bit 2 <-> STM Status/Status/Warning
//     Drive/Inputs/In/nState2 @bit 3 <-> STM Status/Status/Digital input 1
//     Drive/Inputs/In/nState2 @bit 4 <-> STM Status/Status/Digital input 2
//     Drive/Inputs/In/nState2 @bit 5 <-> STM Status/Status/Sync error
//     Drive/Inputs/In/nState2 @bit 7 <-> STM Status/Status/TxPDO Toggle
//     Drive/Inputs/In/nState4 @bit 1 <-> WcState/InputToggle
//     Drive/Inputs/In/nState4 <-> WcState/WcState
//     Drive/Outputs/Out/nCtrl1 <-> STM Control/Control/Enable
//     Drive/Outputs/Out/nCtrl1 @bit 2 <-> STM Control/Control/Reduce torque
//     Drive/Outputs/Out/nCtrl1 @bit 1 <-> STM Control/Control/Reset
//     Drive/Outputs/Out/nDataOut2[0] <-> STM Velocity/Velocity
//   (this object) <-> PLC Rail (EtherCAT)/Power (EK1200)/PLC Junction 2 (EK1122)/X1 HXR EC1 (EK1100)/EC1 E1 (EK1122)/X1 SL1L0-Power (EK1100)/SL1L0-EL5042-E6
//     Enc/Inputs/In/nComState @bit 1 <-> WcState/InputToggle
//     Enc/Inputs/In/nComState <-> WcState/WcState
//     Enc/Inputs/In/nDataIn1 <-> FB Inputs Channel 1/Position
//     Enc/Inputs/In/nDataIn1 <-> FB Inputs Channel 2/Position
//     Enc/Inputs/In/nState1 @bit 12 <-> FB Inputs Channel 1/Status/Diag
//     Enc/Inputs/In/nState1 @bit 12 <-> FB Inputs Channel 2/Status/Diag
//     Enc/Inputs/In/nState1 @bit 1 <-> FB Inputs Channel 1/Status/Error
//     Enc/Inputs/In/nState1 @bit 1 <-> FB Inputs Channel 2/Status/Error
//     Enc/Inputs/In/nState1 @bit 14 <-> FB Inputs Channel 1/Status/Input cycle counter
//     Enc/Inputs/In/nState1 @bit 14 <-> FB Inputs Channel 2/Status/Input cycle counter
//     Enc/Inputs/In/nState1 @bit 2 <-> FB Inputs Channel 1/Status/Ready
//     Enc/Inputs/In/nState1 @bit 2 <-> FB Inputs Channel 2/Status/Ready
//     Enc/Inputs/In/nState1 @bit 13 <-> FB Inputs Channel 1/Status/TxPDO State
//     Enc/Inputs/In/nState1 @bit 13 <-> FB Inputs Channel 2/Status/TxPDO State
//     Enc/Inputs/In/nState1 <-> FB Inputs Channel 1/Status/Warning
//     Enc/Inputs/In/nState1 <-> FB Inputs Channel 2/Status/Warning
//   (this object) <-> PLC Rail (EtherCAT)/Power (EK1200)/PLC Junction 2 (EK1122)/X1 HXR EC1 (EK1100)/EC1 E1 (EK1122)/X1 SL1L0-Power (EK1100)/SL1L0-EL7041-E5
//     Drive/Inputs/In/nState1 @bit 3 <-> STM Status/Status/Error
//     Drive/Inputs/In/nState1 @bit 5 <-> STM Status/Status/Moving negative
//     Drive/Inputs/In/nState1 @bit 4 <-> STM Status/Status/Moving positive
//     Drive/Inputs/In/nState1 @bit 1 <-> STM Status/Status/Ready
//     Drive/Inputs/In/nState1 <-> STM Status/Status/Ready to enable
//     Drive/Inputs/In/nState1 @bit 6 <-> STM Status/Status/Torque reduced
//     Drive/Inputs/In/nState1 @bit 2 <-> STM Status/Status/Warning
//     Drive/Inputs/In/nState2 @bit 3 <-> STM Status/Status/Digital input 1
//     Drive/Inputs/In/nState2 @bit 4 <-> STM Status/Status/Digital input 2
//     Drive/Inputs/In/nState2 @bit 5 <-> STM Status/Status/Sync error
//     Drive/Inputs/In/nState2 @bit 7 <-> STM Status/Status/TxPDO Toggle
//     Drive/Inputs/In/nState4 @bit 1 <-> WcState/InputToggle
//     Drive/Inputs/In/nState4 <-> WcState/WcState
//     Drive/Outputs/Out/nCtrl1 <-> STM Control/Control/Enable
//     Drive/Outputs/Out/nCtrl1 @bit 2 <-> STM Control/Control/Reduce torque
//     Drive/Outputs/Out/nCtrl1 @bit 1 <-> STM Control/Control/Reset
//     Drive/Outputs/Out/nDataOut2[0] <-> STM Velocity/Velocity
//   (this object) <-> PLC Rail (EtherCAT)/Power (EK1200)/PLC Junction 2 (EK1122)/X1 HXR EC1 (EK1100)/EC1 E1 (EK1122)/X1 SL1L0-Power (EK1100)/SL1L0-EL7041-E7
//     Drive/Inputs/In/nState1 @bit 3 <-> STM Status/Status/Error
//     Drive/Inputs/In/nState1 @bit 5 <-> STM Status/Status/Moving negative
//     Drive/Inputs/In/nState1 @bit 4 <-> STM Status/Status/Moving positive
//     Drive/Inputs/In/nState1 @bit 1 <-> STM Status/Status/Ready
//     Drive/Inputs/In/nState1 <-> STM Status/Status/Ready to enable
//     Drive/Inputs/In/nState1 @bit 6 <-> STM Status/Status/Torque reduced
//     Drive/Inputs/In/nState1 @bit 2 <-> STM Status/Status/Warning
//     Drive/Inputs/In/nState2 @bit 3 <-> STM Status/Status/Digital input 1
//     Drive/Inputs/In/nState2 @bit 4 <-> STM Status/Status/Digital input 2
//     Drive/Inputs/In/nState2 @bit 5 <-> STM Status/Status/Sync error
//     Drive/Inputs/In/nState2 @bit 7 <-> STM Status/Status/TxPDO Toggle
//     Drive/Inputs/In/nState4 @bit 1 <-> WcState/InputToggle
//     Drive/Inputs/In/nState4 <-> WcState/WcState
//     Drive/Outputs/Out/nCtrl1 <-> STM Control/Control/Enable
//     Drive/Outputs/Out/nCtrl1 @bit 2 <-> STM Control/Control/Reduce torque
//     Drive/Outputs/Out/nCtrl1 @bit 1 <-> STM Control/Control/Reset
//     Drive/Outputs/Out/nDataOut2[0] <-> STM Velocity/Velocity
//   (this object) <-> PLC Rail (EtherCAT)/Power (EK1200)/PLC Junction 2 (EK1122)/X1 HXR EC1 (EK1100)/EC1 E2 (EK1122)/X2 SL2L0-Power (EK1100)/SL2L0-EL5042-E2
//     Enc/Inputs/In/nComState @bit 1 <-> WcState/InputToggle
//     Enc/Inputs/In/nComState <-> WcState/WcState
//     Enc/Inputs/In/nDataIn1 <-> FB Inputs Channel 1/Position
//     Enc/Inputs/In/nDataIn1 <-> FB Inputs Channel 2/Position
//     Enc/Inputs/In/nState1 @bit 12 <-> FB Inputs Channel 1/Status/Diag
//     Enc/Inputs/In/nState1 @bit 12 <-> FB Inputs Channel 2/Status/Diag
//     Enc/Inputs/In/nState1 @bit 1 <-> FB Inputs Channel 1/Status/Error
//     Enc/Inputs/In/nState1 @bit 1 <-> FB Inputs Channel 2/Status/Error
//     Enc/Inputs/In/nState1 @bit 14 <-> FB Inputs Channel 1/Status/Input cycle counter
//     Enc/Inputs/In/nState1 @bit 14 <-> FB Inputs Channel 2/Status/Input cycle counter
//     Enc/Inputs/In/nState1 @bit 2 <-> FB Inputs Channel 1/Status/Ready
//     Enc/Inputs/In/nState1 @bit 2 <-> FB Inputs Channel 2/Status/Ready
//     Enc/Inputs/In/nState1 @bit 13 <-> FB Inputs Channel 1/Status/TxPDO State
//     Enc/Inputs/In/nState1 @bit 13 <-> FB Inputs Channel 2/Status/TxPDO State
//     Enc/Inputs/In/nState1 <-> FB Inputs Channel 1/Status/Warning
//     Enc/Inputs/In/nState1 <-> FB Inputs Channel 2/Status/Warning
//   (this object) <-> PLC Rail (EtherCAT)/Power (EK1200)/PLC Junction 2 (EK1122)/X1 HXR EC1 (EK1100)/EC1 E2 (EK1122)/X2 SL2L0-Power (EK1100)/SL2L0-EL7041-E1
//     Drive/Inputs/In/nState1 @bit 3 <-> STM Status/Status/Error
//     Drive/Inputs/In/nState1 @bit 5 <-> STM Status/Status/Moving negative
//     Drive/Inputs/In/nState1 @bit 4 <-> STM Status/Status/Moving positive
//     Drive/Inputs/In/nState1 @bit 1 <-> STM Status/Status/Ready
//     Drive/Inputs/In/nState1 <-> STM Status/Status/Ready to enable
//     Drive/Inputs/In/nState1 @bit 6 <-> STM Status/Status/Torque reduced
//     Drive/Inputs/In/nState1 @bit 2 <-> STM Status/Status/Warning
//     Drive/Inputs/In/nState2 @bit 3 <-> STM Status/Status/Digital input 1
//     Drive/Inputs/In/nState2 @bit 4 <-> STM Status/Status/Digital input 2
//     Drive/Inputs/In/nState2 @bit 5 <-> STM Status/Status/Sync error
//     Drive/Inputs/In/nState2 @bit 7 <-> STM Status/Status/TxPDO Toggle
//     Drive/Inputs/In/nState4 @bit 1 <-> WcState/InputToggle
//     Drive/Inputs/In/nState4 <-> WcState/WcState
//     Drive/Outputs/Out/nCtrl1 <-> STM Control/Control/Enable
//     Drive/Outputs/Out/nCtrl1 @bit 2 <-> STM Control/Control/Reduce torque
//     Drive/Outputs/Out/nCtrl1 @bit 1 <-> STM Control/Control/Reset
//     Drive/Outputs/Out/nDataOut2[0] <-> STM Velocity/Velocity
//   (this object) <-> PLC Rail (EtherCAT)/Power (EK1200)/PLC Junction 2 (EK1122)/X1 HXR EC1 (EK1100)/EC1 E2 (EK1122)/X2 SL2L0-Power (EK1100)/SL2L0-EL7041-E3
//     Drive/Inputs/In/nState1 @bit 3 <-> STM Status/Status/Error
//     Drive/Inputs/In/nState1 @bit 5 <-> STM Status/Status/Moving negative
//     Drive/Inputs/In/nState1 @bit 4 <-> STM Status/Status/Moving positive
//     Drive/Inputs/In/nState1 @bit 1 <-> STM Status/Status/Ready
//     Drive/Inputs/In/nState1 <-> STM Status/Status/Ready to enable
//     Drive/Inputs/In/nState1 @bit 6 <-> STM Status/Status/Torque reduced
//     Drive/Inputs/In/nState1 @bit 2 <-> STM Status/Status/Warning
//     Drive/Inputs/In/nState2 @bit 3 <-> STM Status/Status/Digital input 1
//     Drive/Inputs/In/nState2 @bit 4 <-> STM Status/Status/Digital input 2
//     Drive/Inputs/In/nState2 @bit 5 <-> STM Status/Status/Sync error
//     Drive/Inputs/In/nState2 @bit 7 <-> STM Status/Status/TxPDO Toggle
//     Drive/Inputs/In/nState4 @bit 1 <-> WcState/InputToggle
//     Drive/Inputs/In/nState4 <-> WcState/WcState
//     Drive/Outputs/Out/nCtrl1 <-> STM Control/Control/Enable
//     Drive/Outputs/Out/nCtrl1 @bit 2 <-> STM Control/Control/Reduce torque
//     Drive/Outputs/Out/nCtrl1 @bit 1 <-> STM Control/Control/Reset
//     Drive/Outputs/Out/nDataOut2[0] <-> STM Velocity/Velocity
//   (this object) <-> PLC Rail (EtherCAT)/Power (EK1200)/PLC Junction 2 (EK1122)/X1 HXR EC1 (EK1100)/EC1 E2 (EK1122)/X2 SL2L0-Power (EK1100)/SL2L0-EL5042-E6
//     Enc/Inputs/In/nComState @bit 1 <-> WcState/InputToggle
//     Enc/Inputs/In/nComState <-> WcState/WcState
//     Enc/Inputs/In/nDataIn1 <-> FB Inputs Channel 1/Position
//     Enc/Inputs/In/nDataIn1 <-> FB Inputs Channel 2/Position
//     Enc/Inputs/In/nState1 @bit 12 <-> FB Inputs Channel 1/Status/Diag
//     Enc/Inputs/In/nState1 @bit 12 <-> FB Inputs Channel 2/Status/Diag
//     Enc/Inputs/In/nState1 @bit 1 <-> FB Inputs Channel 1/Status/Error
//     Enc/Inputs/In/nState1 @bit 1 <-> FB Inputs Channel 2/Status/Error
//     Enc/Inputs/In/nState1 @bit 14 <-> FB Inputs Channel 1/Status/Input cycle counter
//     Enc/Inputs/In/nState1 @bit 14 <-> FB Inputs Channel 2/Status/Input cycle counter
//     Enc/Inputs/In/nState1 @bit 2 <-> FB Inputs Channel 1/Status/Ready
//     Enc/Inputs/In/nState1 @bit 2 <-> FB Inputs Channel 2/Status/Ready
//     Enc/Inputs/In/nState1 @bit 13 <-> FB Inputs Channel 1/Status/TxPDO State
//     Enc/Inputs/In/nState1 @bit 13 <-> FB Inputs Channel 2/Status/TxPDO State
//     Enc/Inputs/In/nState1 <-> FB Inputs Channel 1/Status/Warning
//     Enc/Inputs/In/nState1 <-> FB Inputs Channel 2/Status/Warning
//   (this object) <-> PLC Rail (EtherCAT)/Power (EK1200)/PLC Junction 2 (EK1122)/X1 HXR EC1 (EK1100)/EC1 E2 (EK1122)/X2 SL2L0-Power (EK1100)/SL2L0-EL7041-E5
//     Drive/Inputs/In/nState1 @bit 3 <-> STM Status/Status/Error
//     Drive/Inputs/In/nState1 @bit 5 <-> STM Status/Status/Moving negative
//     Drive/Inputs/In/nState1 @bit 4 <-> STM Status/Status/Moving positive
//     Drive/Inputs/In/nState1 @bit 1 <-> STM Status/Status/Ready
//     Drive/Inputs/In/nState1 <-> STM Status/Status/Ready to enable
//     Drive/Inputs/In/nState1 @bit 6 <-> STM Status/Status/Torque reduced
//     Drive/Inputs/In/nState1 @bit 2 <-> STM Status/Status/Warning
//     Drive/Inputs/In/nState2 @bit 3 <-> STM Status/Status/Digital input 1
//     Drive/Inputs/In/nState2 @bit 4 <-> STM Status/Status/Digital input 2
//     Drive/Inputs/In/nState2 @bit 5 <-> STM Status/Status/Sync error
//     Drive/Inputs/In/nState2 @bit 7 <-> STM Status/Status/TxPDO Toggle
//     Drive/Inputs/In/nState4 @bit 1 <-> WcState/InputToggle
//     Drive/Inputs/In/nState4 <-> WcState/WcState
//     Drive/Outputs/Out/nCtrl1 <-> STM Control/Control/Enable
//     Drive/Outputs/Out/nCtrl1 @bit 2 <-> STM Control/Control/Reduce torque
//     Drive/Outputs/Out/nCtrl1 @bit 1 <-> STM Control/Control/Reset
//     Drive/Outputs/Out/nDataOut2[0] <-> STM Velocity/Velocity
//   (this object) <-> PLC Rail (EtherCAT)/Power (EK1200)/PLC Junction 2 (EK1122)/X1 HXR EC1 (EK1100)/EC1 E2 (EK1122)/X2 SL2L0-Power (EK1100)/SL2L0-EL7041-E7
//     Drive/Inputs/In/nState1 @bit 3 <-> STM Status/Status/Error
//     Drive/Inputs/In/nState1 @bit 5 <-> STM Status/Status/Moving negative
//     Drive/Inputs/In/nState1 @bit 4 <-> STM Status/Status/Moving positive
//     Drive/Inputs/In/nState1 @bit 1 <-> STM Status/Status/Ready
//     Drive/Inputs/In/nState1 <-> STM Status/Status/Ready to enable
//     Drive/Inputs/In/nState1 @bit 6 <-> STM Status/Status/Torque reduced
//     Drive/Inputs/In/nState1 @bit 2 <-> STM Status/Status/Warning
//     Drive/Inputs/In/nState2 @bit 3 <-> STM Status/Status/Digital input 1
//     Drive/Inputs/In/nState2 @bit 4 <-> STM Status/Status/Digital input 2
//     Drive/Inputs/In/nState2 @bit 5 <-> STM Status/Status/Sync error
//     Drive/Inputs/In/nState2 @bit 7 <-> STM Status/Status/TxPDO Toggle
//     Drive/Inputs/In/nState4 @bit 1 <-> WcState/InputToggle
//     Drive/Inputs/In/nState4 <-> WcState/WcState
//     Drive/Outputs/Out/nCtrl1 <-> STM Control/Control/Enable
//     Drive/Outputs/Out/nCtrl1 @bit 2 <-> STM Control/Control/Reduce torque
//     Drive/Outputs/Out/nCtrl1 @bit 1 <-> STM Control/Control/Reset
//     Drive/Outputs/Out/nDataOut2[0] <-> STM Velocity/Velocity
//   (this object) <-> PLC Rail (EtherCAT)/Power (EK1200)/PLC Junction 2 (EK1122)/X1 HXR EC1 (EK1100)/EC1 E3 (EK1122)/X2_0 SP1L0-KMONO_MOTOR (EK1100)/SP1L0-EL7031-E1-MOTORS
//     Drive/Inputs/In/nState1 @bit 3 <-> STM Status/Status/Error
//     Drive/Inputs/In/nState1 @bit 5 <-> STM Status/Status/Moving negative
//     Drive/Inputs/In/nState1 @bit 4 <-> STM Status/Status/Moving positive
//     Drive/Inputs/In/nState1 @bit 1 <-> STM Status/Status/Ready
//     Drive/Inputs/In/nState1 <-> STM Status/Status/Ready to enable
//     Drive/Inputs/In/nState1 @bit 6 <-> STM Status/Status/Torque reduced
//     Drive/Inputs/In/nState1 @bit 2 <-> STM Status/Status/Warning
//     Drive/Inputs/In/nState2 @bit 3 <-> STM Status/Status/Digital input 1
//     Drive/Inputs/In/nState2 @bit 4 <-> STM Status/Status/Digital input 2
//     Drive/Inputs/In/nState2 @bit 5 <-> STM Status/Status/Sync error
//     Drive/Inputs/In/nState2 @bit 7 <-> STM Status/Status/TxPDO Toggle
//     Drive/Inputs/In/nState4 @bit 1 <-> WcState/InputToggle
//     Drive/Inputs/In/nState4 <-> WcState/WcState
//     Drive/Outputs/Out/nCtrl1 <-> STM Control/Control/Enable
//     Drive/Outputs/Out/nCtrl1 @bit 2 <-> STM Control/Control/Reduce torque
//     Drive/Outputs/Out/nCtrl1 @bit 1 <-> STM Control/Control/Reset
//     Drive/Outputs/Out/nDataOut2[0] <-> STM Velocity/Velocity
//     Enc/Inputs/In/nDataIn1[0] <-> ENC Status compact/Counter value
//     Enc/Inputs/In/nDataIn2[0] <-> ENC Status compact/Latch value
//     Enc/Inputs/In/nState1 @bit 4 <-> ENC Status compact/Status/Counter overflow
//     Enc/Inputs/In/nState1 @bit 3 <-> ENC Status compact/Status/Counter underflow
//     Enc/Inputs/In/nState1 @bit 1 <-> ENC Status compact/Status/Latch extern valid
//     Enc/Inputs/In/nState1 @bit 2 <-> ENC Status compact/Status/Set counter done
//     Enc/Inputs/In/nState2 @bit 4 <-> ENC Status compact/Status/Status of extern latch
//     Enc/Inputs/In/nState2 @bit 5 <-> ENC Status compact/Status/Sync error
//     Enc/Inputs/In/nState2 @bit 7 <-> ENC Status compact/Status/TxPDO Toggle
//     Enc/Inputs/In/nState4 @bit 1 <-> WcState/InputToggle
//     Enc/Inputs/In/nState4 <-> WcState/WcState
//     Enc/Outputs/Out/nCtrl1 @bit 3 <-> ENC Control compact/Control/Enable latch extern on negative edge
//     Enc/Outputs/Out/nCtrl1 @bit 1 <-> ENC Control compact/Control/Enable latch extern on positive edge
//     Enc/Outputs/Out/nCtrl1 @bit 2 <-> ENC Control compact/Control/Set counter
//     Enc/Outputs/Out/nDataOut1[0] <-> ENC Control compact/Set counter value
//   (this object) <-> PLC Rail (EtherCAT)/Power (EK1200)/PLC Junction 2 (EK1122)/X1 HXR EC1 (EK1100)/EC1 E3 (EK1122)/X2_0 SP1L0-KMONO_MOTOR (EK1100)/SP1L0-EL7041-E2-MOTORS
//     Drive/Inputs/In/nState1 @bit 3 <-> STM Status/Status/Error
//     Drive/Inputs/In/nState1 @bit 5 <-> STM Status/Status/Moving negative
//     Drive/Inputs/In/nState1 @bit 4 <-> STM Status/Status/Moving positive
//     Drive/Inputs/In/nState1 @bit 1 <-> STM Status/Status/Ready
//     Drive/Inputs/In/nState1 <-> STM Status/Status/Ready to enable
//     Drive/Inputs/In/nState1 @bit 6 <-> STM Status/Status/Torque reduced
//     Drive/Inputs/In/nState1 @bit 2 <-> STM Status/Status/Warning
//     Drive/Inputs/In/nState2 @bit 3 <-> STM Status/Status/Digital input 1
//     Drive/Inputs/In/nState2 @bit 4 <-> STM Status/Status/Digital input 2
//     Drive/Inputs/In/nState2 @bit 5 <-> STM Status/Status/Sync error
//     Drive/Inputs/In/nState2 @bit 7 <-> STM Status/Status/TxPDO Toggle
//     Drive/Inputs/In/nState4 @bit 1 <-> WcState/InputToggle
//     Drive/Inputs/In/nState4 <-> WcState/WcState
//     Drive/Outputs/Out/nCtrl1 <-> STM Control/Control/Enable
//     Drive/Outputs/Out/nCtrl1 @bit 2 <-> STM Control/Control/Reduce torque
//     Drive/Outputs/Out/nCtrl1 @bit 1 <-> STM Control/Control/Reset
//     Drive/Outputs/Out/nDataOut2[0] <-> STM Velocity/Velocity
//   (this object) <-> PLC Rail (EtherCAT)/Power (EK1200)/PLC Junction 2 (EK1122)/X1 HXR EC1 (EK1100)/EC1 E3 (EK1122)/X2_1 SP1L0-KMONO_LVDT (EK1100)/SP1L0-EL3052-E4-LVDT
//     Enc/Inputs/In/nDataIn1[0] <-> AI Standard Channel 1/Value
//     Enc/Inputs/In/nDataIn1[0] <-> AI Standard Channel 2/Value
//     Enc/Inputs/In/nState4 @bit 1 <-> WcState/InputToggle
//     Enc/Inputs/In/nState4 <-> WcState/WcState
//   (this object) <-> PLC Rail (EtherCAT)/Power (EK1200)/PLC Junction 2 (EK1122)/X1 HXR EC1 (EK1100)/EC1 E3 (EK1122)/X2_0 SP1L0-KMONO_MOTOR (EK1100)/SP1L0-EL7041-E3-MOTORS
//     Drive/Inputs/In/nState1 @bit 3 <-> STM Status/Status/Error
//     Drive/Inputs/In/nState1 @bit 5 <-> STM Status/Status/Moving negative
//     Drive/Inputs/In/nState1 @bit 4 <-> STM Status/Status/Moving positive
//     Drive/Inputs/In/nState1 @bit 1 <-> STM Status/Status/Ready
//     Drive/Inputs/In/nState1 <-> STM Status/Status/Ready to enable
//     Drive/Inputs/In/nState1 @bit 6 <-> STM Status/Status/Torque reduced
//     Drive/Inputs/In/nState1 @bit 2 <-> STM Status/Status/Warning
//     Drive/Inputs/In/nState2 @bit 3 <-> STM Status/Status/Digital input 1
//     Drive/Inputs/In/nState2 @bit 4 <-> STM Status/Status/Digital input 2
//     Drive/Inputs/In/nState2 @bit 5 <-> STM Status/Status/Sync error
//     Drive/Inputs/In/nState2 @bit 7 <-> STM Status/Status/TxPDO Toggle
//     Drive/Inputs/In/nState4 @bit 1 <-> WcState/InputToggle
//     Drive/Inputs/In/nState4 <-> WcState/WcState
//     Drive/Outputs/Out/nCtrl1 <-> STM Control/Control/Enable
//     Drive/Outputs/Out/nCtrl1 @bit 2 <-> STM Control/Control/Reduce torque
//     Drive/Outputs/Out/nCtrl1 @bit 1 <-> STM Control/Control/Reset
//     Drive/Outputs/Out/nDataOut2[0] <-> STM Velocity/Velocity
//   (this object) <-> PLC Rail (EtherCAT)/Power (EK1200)/PLC Junction 2 (EK1122)/X1 HXR EC1 (EK1100)/EC1 E3 (EK1122)/X2_0 SP1L0-KMONO_MOTOR (EK1100)/SP1L0-EL7041-E4-MOTORS
//     Drive/Inputs/In/nState1 @bit 3 <-> STM Status/Status/Error
//     Drive/Inputs/In/nState1 @bit 5 <-> STM Status/Status/Moving negative
//     Drive/Inputs/In/nState1 @bit 4 <-> STM Status/Status/Moving positive
//     Drive/Inputs/In/nState1 @bit 1 <-> STM Status/Status/Ready
//     Drive/Inputs/In/nState1 <-> STM Status/Status/Ready to enable
//     Drive/Inputs/In/nState1 @bit 6 <-> STM Status/Status/Torque reduced
//     Drive/Inputs/In/nState1 @bit 2 <-> STM Status/Status/Warning
//     Drive/Inputs/In/nState2 @bit 3 <-> STM Status/Status/Digital input 1
//     Drive/Inputs/In/nState2 @bit 4 <-> STM Status/Status/Digital input 2
//     Drive/Inputs/In/nState2 @bit 5 <-> STM Status/Status/Sync error
//     Drive/Inputs/In/nState2 @bit 7 <-> STM Status/Status/TxPDO Toggle
//     Drive/Inputs/In/nState4 @bit 1 <-> WcState/InputToggle
//     Drive/Inputs/In/nState4 <-> WcState/WcState
//     Drive/Outputs/Out/nCtrl1 <-> STM Control/Control/Enable
//     Drive/Outputs/Out/nCtrl1 @bit 2 <-> STM Control/Control/Reduce torque
//     Drive/Outputs/Out/nCtrl1 @bit 1 <-> STM Control/Control/Reset
//     Drive/Outputs/Out/nDataOut2[0] <-> STM Velocity/Velocity
//     Enc/Inputs/In/nDataIn1[0] <-> ENC Status compact/Counter value
//     Enc/Inputs/In/nDataIn2[0] <-> ENC Status compact/Latch value
//     Enc/Inputs/In/nState1 @bit 4 <-> ENC Status compact/Status/Counter overflow
//     Enc/Inputs/In/nState1 @bit 3 <-> ENC Status compact/Status/Counter underflow
//     Enc/Inputs/In/nState1 @bit 7 <-> ENC Status compact/Status/Extrapolation stall
//     Enc/Inputs/In/nState1 <-> ENC Status compact/Status/Latch C valid
//     Enc/Inputs/In/nState1 @bit 1 <-> ENC Status compact/Status/Latch extern valid
//     Enc/Inputs/In/nState1 @bit 2 <-> ENC Status compact/Status/Set counter done
//     Enc/Inputs/In/nState2 @bit 4 <-> ENC Status compact/Status/Status of extern latch
//     Enc/Inputs/In/nState2 <-> ENC Status compact/Status/Status of input A
//     Enc/Inputs/In/nState2 @bit 1 <-> ENC Status compact/Status/Status of input B
//     Enc/Inputs/In/nState2 @bit 2 <-> ENC Status compact/Status/Status of input C
//     Enc/Inputs/In/nState2 @bit 5 <-> ENC Status compact/Status/Sync error
//     Enc/Inputs/In/nState2 @bit 7 <-> ENC Status compact/Status/TxPDO Toggle
//     Enc/Inputs/In/nState4 @bit 1 <-> WcState/InputToggle
//     Enc/Inputs/In/nState4 <-> WcState/WcState
//     Enc/Outputs/Out/nCtrl1 <-> ENC Control compact/Control/Enable latch C
//     Enc/Outputs/Out/nCtrl1 @bit 3 <-> ENC Control compact/Control/Enable latch extern on negative edge
//     Enc/Outputs/Out/nCtrl1 @bit 1 <-> ENC Control compact/Control/Enable latch extern on positive edge
//     Enc/Outputs/Out/nCtrl1 @bit 2 <-> ENC Control compact/Control/Set counter
//     Enc/Outputs/Out/nDataOut1[0] <-> ENC Control compact/Set counter value
//   (this object) <-> PLC Rail (EtherCAT)/Power (EK1200)/PLC Junction 2 (EK1122)/X1 HXR EC1 (EK1100)/EC1 E3 (EK1122)/X2_0 SP1L0-KMONO_MOTOR (EK1100)/SP1L0-EL7041-E5-MOTORS
//     Drive/Inputs/In/nState1 @bit 3 <-> STM Status/Status/Error
//     Drive/Inputs/In/nState1 @bit 5 <-> STM Status/Status/Moving negative
//     Drive/Inputs/In/nState1 @bit 4 <-> STM Status/Status/Moving positive
//     Drive/Inputs/In/nState1 @bit 1 <-> STM Status/Status/Ready
//     Drive/Inputs/In/nState1 <-> STM Status/Status/Ready to enable
//     Drive/Inputs/In/nState1 @bit 6 <-> STM Status/Status/Torque reduced
//     Drive/Inputs/In/nState1 @bit 2 <-> STM Status/Status/Warning
//     Drive/Inputs/In/nState2 @bit 3 <-> STM Status/Status/Digital input 1
//     Drive/Inputs/In/nState2 @bit 4 <-> STM Status/Status/Digital input 2
//     Drive/Inputs/In/nState2 @bit 5 <-> STM Status/Status/Sync error
//     Drive/Inputs/In/nState2 @bit 7 <-> STM Status/Status/TxPDO Toggle
//     Drive/Inputs/In/nState4 @bit 1 <-> WcState/InputToggle
//     Drive/Inputs/In/nState4 <-> WcState/WcState
//     Drive/Outputs/Out/nCtrl1 <-> STM Control/Control/Enable
//     Drive/Outputs/Out/nCtrl1 @bit 2 <-> STM Control/Control/Reduce torque
//     Drive/Outputs/Out/nCtrl1 @bit 1 <-> STM Control/Control/Reset
//     Drive/Outputs/Out/nDataOut2[0] <-> STM Velocity/Velocity
//   (this object) <-> PLC Rail (EtherCAT)/Power (EK1200)/PLC Junction 2 (EK1122)/X1 HXR EC1 (EK1100)/EC1 E3 (EK1122)/X2_1 SP1L0-KMONO_LVDT (EK1100)/SP1L0-EL3052-E5-LVDT
//     Enc/Inputs/In/nDataIn1[0] <-> AI Standard Channel 2/Value
//     Enc/Inputs/In/nState4 @bit 1 <-> WcState/InputToggle
//     Enc/Inputs/In/nState4 <-> WcState/WcState
//   (this object) <-> PLC Rail (EtherCAT)/Power (EK1200)/PLC Junction 2 (EK1122)/X1 HXR EC1 (EK1100)/EC1 E3 (EK1122)/X2_0 SP1L0-KMONO_MOTOR (EK1100)/SP1L0-EL7041-E6-MOTORS
//     Drive/Inputs/In/nState1 @bit 3 <-> STM Status/Status/Error
//     Drive/Inputs/In/nState1 @bit 5 <-> STM Status/Status/Moving negative
//     Drive/Inputs/In/nState1 @bit 4 <-> STM Status/Status/Moving positive
//     Drive/Inputs/In/nState1 @bit 1 <-> STM Status/Status/Ready
//     Drive/Inputs/In/nState1 <-> STM Status/Status/Ready to enable
//     Drive/Inputs/In/nState1 @bit 6 <-> STM Status/Status/Torque reduced
//     Drive/Inputs/In/nState1 @bit 2 <-> STM Status/Status/Warning
//     Drive/Inputs/In/nState2 @bit 3 <-> STM Status/Status/Digital input 1
//     Drive/Inputs/In/nState2 @bit 4 <-> STM Status/Status/Digital input 2
//     Drive/Inputs/In/nState2 @bit 5 <-> STM Status/Status/Sync error
//     Drive/Inputs/In/nState2 @bit 7 <-> STM Status/Status/TxPDO Toggle
//     Drive/Inputs/In/nState4 @bit 1 <-> WcState/InputToggle
//     Drive/Inputs/In/nState4 <-> WcState/WcState
//     Drive/Outputs/Out/nCtrl1 <-> STM Control/Control/Enable
//     Drive/Outputs/Out/nCtrl1 @bit 2 <-> STM Control/Control/Reduce torque
//     Drive/Outputs/Out/nCtrl1 @bit 1 <-> STM Control/Control/Reset
//     Drive/Outputs/Out/nDataOut2[0] <-> STM Velocity/Velocity
//   (this object) <-> PLC Rail (EtherCAT)/Power (EK1200)/PLC Junction 2 (EK1122)/X1 HXR EC1 (EK1100)/EC1 E3 (EK1122)/X2_1 SP1L0-KMONO_LVDT (EK1100)/SP1L0-EL3052-E6-LVDT
//     Enc/Inputs/In/nDataIn1[0] <-> AI Standard Channel 1/Value
//     Enc/Inputs/In/nState4 @bit 1 <-> WcState/InputToggle
//     Enc/Inputs/In/nState4 <-> WcState/WcState
//   lfe_motion Instance <-> PLC Rail (EtherCAT)/Power (EK1200)/PLC Junction 1 (EK1122)/X1 RTDSL0 (EK1100)/RTDSL0-EL7041-01
//     PlcTask Inputs/Main.M33.bLimitBackwardEnable <-> STM Status/Status/Digital input 2
//     PlcTask Inputs/Main.M33.bLimitForwardEnable <-> STM Status/Status/Digital input 1
//   lfe_motion Instance <-> PLC Rail (EtherCAT)/Power (EK1200)/PLC Junction 1 (EK1122)/X1 RTDSL0 (EK1100)/RTDSL0-EL7041-05
//     PlcTask Inputs/Main.M38.bLimitBackwardEnable <-> STM Status/Status/Digital input 2
//     PlcTask Inputs/Main.M38.bLimitForwardEnable <-> STM Status/Status/Digital input 1
//   lfe_motion Instance <-> PLC Rail (EtherCAT)/Power (EK1200)/PLC Junction 1 (EK1122)/X1 RTDSL0 (EK1100)/RTDSL0-MPA-EL1008
//     PlcTask Inputs/RTDSL0.RTDSL0_MPA_01.i_xInsertedLS <-> Channel 1/Input
//     PlcTask Inputs/RTDSL0.RTDSL0_MPA_02.i_xInsertedLS <-> Channel 3/Input
//     PlcTask Inputs/RTDSL0.RTDSL0_MPA_03.i_xInsertedLS <-> Channel 5/Input
//     PlcTask Inputs/RTDSL0.RTDSL0_MPA_04.i_xInsertedLS <-> Channel 7/Input
//     PlcTask Inputs/RTDSL0.RTDSL0_MPA_01.i_xRetractedLS <-> Channel 2/Input
//     PlcTask Inputs/RTDSL0.RTDSL0_MPA_02.i_xRetractedLS <-> Channel 4/Input
//     PlcTask Inputs/RTDSL0.RTDSL0_MPA_03.i_xRetractedLS <-> Channel 6/Input
//     PlcTask Inputs/RTDSL0.RTDSL0_MPA_04.i_xRetractedLS <-> Channel 8/Input
//   lfe_motion Instance <-> PLC Rail (EtherCAT)/Power (EK1200)/PLC Junction 1 (EK1122)/X1 RTDSL0 (EK1100)/RTDSL0-MPA-EL2008
//     PlcTask Outputs/RTDSL0.RTDSL0_MPA_01.q_xInsert_DO <-> Channel 1/Output
//     PlcTask Outputs/RTDSL0.RTDSL0_MPA_02.q_xInsert_DO <-> Channel 3/Output
//     PlcTask Outputs/RTDSL0.RTDSL0_MPA_03.q_xInsert_DO <-> Channel 5/Output
//     PlcTask Outputs/RTDSL0.RTDSL0_MPA_04.q_xInsert_DO <-> Channel 7/Output
//     PlcTask Outputs/RTDSL0.RTDSL0_MPA_01.q_xRetract_DO <-> Channel 2/Output
//     PlcTask Outputs/RTDSL0.RTDSL0_MPA_02.q_xRetract_DO <-> Channel 4/Output
//     PlcTask Outputs/RTDSL0.RTDSL0_MPA_03.q_xRetract_DO <-> Channel 6/Output
//     PlcTask Outputs/RTDSL0.RTDSL0_MPA_04.q_xRetract_DO <-> Channel 8/Output
//   lfe_motion Instance <-> PLC Rail (EtherCAT)/Power (EK1200)/PLC Junction 1 (EK1122)/X1 RTDSL0 (EK1100)/Term 113 (EL3054)
//     PlcTask Inputs/Main.M38.nRawEncoderINT <-> AI Standard Channel 1/Value
//   lfe_motion Instance <-> PLC Rail (EtherCAT)/Power (EK1200)/PLC Junction 1 (EK1122)/X2 IM1L0-XTES (EK1100)/IM1L0-EL1088
//     PlcTask Inputs/Main.M21.bHome <-> Channel 2/Input
//     PlcTask Inputs/Main.M22.bHome <-> Channel 4/Input
//     PlcTask Inputs/PRG_IM1L0_XTES.fbIM1L0.bFocusEndBwd <-> Channel 4/Input
//     PlcTask Inputs/PRG_IM1L0_XTES.fbIM1L0.bFocusEndFwd <-> Channel 3/Input
//     PlcTask Inputs/PRG_IM1L0_XTES.fbIM1L0.bZoomEndBwd <-> Channel 2/Input
//     PlcTask Inputs/PRG_IM1L0_XTES.fbIM1L0.bZoomEndFwd <-> Channel 1/Input
//   lfe_motion Instance <-> PLC Rail (EtherCAT)/Power (EK1200)/PLC Junction 1 (EK1122)/X2 IM1L0-XTES (EK1100)/IM1L0-EL2004
//     PlcTask Outputs/Main.M20.bBrakeRelease <-> Channel 1/Output
//     PlcTask Outputs/PRG_IM1L0_XTES.fbIM1L0.fbLED.bLEDPower <-> Channel 3/Output
//     PlcTask Outputs/PRG_IM1L0_XTES.fbIM1L0.fbOpal.bOpalPower <-> Channel 2/Output
//   lfe_motion Instance <-> PLC Rail (EtherCAT)/Power (EK1200)/PLC Junction 1 (EK1122)/X2 IM1L0-XTES (EK1100)/IM1L0-EL6002
//     PlcTask Inputs/PRG_IM1L0_XTES.stEL6In/D[{0..21}] <-> COM TxPDO-Map Inputs Channel 1/Data In {0..21}  (22 links)
//     PlcTask Inputs/PRG_IM1L0_XTES.stEL6In/Status <-> COM TxPDO-Map Inputs Channel 1/Status
//     PlcTask Outputs/PRG_IM1L0_XTES.stEL6Out/Ctrl <-> COM RxPDO-Map Outputs Channel 1/Ctrl
//     PlcTask Outputs/PRG_IM1L0_XTES.stEL6Out/D[{0..21}] <-> COM RxPDO-Map Outputs Channel 1/Data Out {0..21}  (22 links)
//   lfe_motion Instance <-> PLC Rail (EtherCAT)/Power (EK1200)/PLC Junction 1 (EK1122)/X2 IM1L0-XTES (EK1100)/IM1L0-EL7041
//     PlcTask Inputs/Main.M20.bLimitForwardEnable <-> STM Status/Status/Digital input 1
//   lfe_motion Instance <-> PLC Rail (EtherCAT)/Power (EK1200)/PLC Junction 2 (EK1122)/X1 HXR EC1 (EK1100)/EC1 E1 (EK1122)/X1 SL1L0-Power (EK1100)/SL1L0-EL3202-E10
//     PlcTask Inputs/PRG_SL1L0_POWER.fbSL1L0.RTD_TOP_1.bError <-> RTD Inputs Channel 1/Status/Error
//     PlcTask Inputs/PRG_SL1L0_POWER.fbSL1L0.RTD_TOP_2.bError <-> RTD Inputs Channel 2/Status/Error
//     PlcTask Inputs/PRG_SL1L0_POWER.fbSL1L0.RTD_TOP_1.bOverrange <-> RTD Inputs Channel 1/Status/Overrange
//     PlcTask Inputs/PRG_SL1L0_POWER.fbSL1L0.RTD_TOP_2.bOverrange <-> RTD Inputs Channel 2/Status/Overrange
//     PlcTask Inputs/PRG_SL1L0_POWER.fbSL1L0.RTD_TOP_1.bUnderrange <-> RTD Inputs Channel 1/Status/Underrange
//     PlcTask Inputs/PRG_SL1L0_POWER.fbSL1L0.RTD_TOP_2.bUnderrange <-> RTD Inputs Channel 2/Status/Underrange
//     PlcTask Inputs/PRG_SL1L0_POWER.fbSL1L0.RTD_TOP_1.iRaw <-> RTD Inputs Channel 1/Value
//     PlcTask Inputs/PRG_SL1L0_POWER.fbSL1L0.RTD_TOP_2.iRaw <-> RTD Inputs Channel 2/Value
//   lfe_motion Instance <-> PLC Rail (EtherCAT)/Power (EK1200)/PLC Junction 2 (EK1122)/X1 HXR EC1 (EK1100)/EC1 E1 (EK1122)/X1 SL1L0-Power (EK1100)/SL1L0-EL3202-E11
//     PlcTask Inputs/PRG_SL1L0_POWER.fbSL1L0.RTD_North_1.bError <-> RTD Inputs Channel 1/Status/Error
//     PlcTask Inputs/PRG_SL1L0_POWER.fbSL1L0.RTD_North_2.bError <-> RTD Inputs Channel 2/Status/Error
//     PlcTask Inputs/PRG_SL1L0_POWER.fbSL1L0.RTD_North_1.bOverrange <-> RTD Inputs Channel 1/Status/Overrange
//     PlcTask Inputs/PRG_SL1L0_POWER.fbSL1L0.RTD_North_2.bOverrange <-> RTD Inputs Channel 2/Status/Overrange
//     PlcTask Inputs/PRG_SL1L0_POWER.fbSL1L0.RTD_North_1.bUnderrange <-> RTD Inputs Channel 1/Status/Underrange
//     PlcTask Inputs/PRG_SL1L0_POWER.fbSL1L0.RTD_North_2.bUnderrange <-> RTD Inputs Channel 2/Status/Underrange
//     PlcTask Inputs/PRG_SL1L0_POWER.fbSL1L0.RTD_North_1.iRaw <-> RTD Inputs Channel 1/Value
//     PlcTask Inputs/PRG_SL1L0_POWER.fbSL1L0.RTD_North_2.iRaw <-> RTD Inputs Channel 2/Value
//   lfe_motion Instance <-> PLC Rail (EtherCAT)/Power (EK1200)/PLC Junction 2 (EK1122)/X1 HXR EC1 (EK1100)/EC1 E1 (EK1122)/X1 SL1L0-Power (EK1100)/SL1L0-EL3202-E8
//     PlcTask Inputs/PRG_SL1L0_POWER.fbSL1L0.RTD_Bottom_1.bError <-> RTD Inputs Channel 1/Status/Error
//     PlcTask Inputs/PRG_SL1L0_POWER.fbSL1L0.RTD_Bottom_2.bError <-> RTD Inputs Channel 2/Status/Error
//     PlcTask Inputs/PRG_SL1L0_POWER.fbSL1L0.RTD_Bottom_1.bOverrange <-> RTD Inputs Channel 1/Status/Overrange
//     PlcTask Inputs/PRG_SL1L0_POWER.fbSL1L0.RTD_Bottom_2.bOverrange <-> RTD Inputs Channel 2/Status/Overrange
//     PlcTask Inputs/PRG_SL1L0_POWER.fbSL1L0.RTD_Bottom_1.bUnderrange <-> RTD Inputs Channel 1/Status/Underrange
//     PlcTask Inputs/PRG_SL1L0_POWER.fbSL1L0.RTD_Bottom_2.bUnderrange <-> RTD Inputs Channel 2/Status/Underrange
//     PlcTask Inputs/PRG_SL1L0_POWER.fbSL1L0.RTD_Bottom_1.iRaw <-> RTD Inputs Channel 1/Value
//     PlcTask Inputs/PRG_SL1L0_POWER.fbSL1L0.RTD_Bottom_2.iRaw <-> RTD Inputs Channel 2/Value
//   lfe_motion Instance <-> PLC Rail (EtherCAT)/Power (EK1200)/PLC Junction 2 (EK1122)/X1 HXR EC1 (EK1100)/EC1 E1 (EK1122)/X1 SL1L0-Power (EK1100)/SL1L0-EL3202-E9
//     PlcTask Inputs/PRG_SL1L0_POWER.fbSL1L0.RTD_South_1.bError <-> RTD Inputs Channel 1/Status/Error
//     PlcTask Inputs/PRG_SL1L0_POWER.fbSL1L0.RTD_South_2.bError <-> RTD Inputs Channel 2/Status/Error
//     PlcTask Inputs/PRG_SL1L0_POWER.fbSL1L0.RTD_South_1.bOverrange <-> RTD Inputs Channel 1/Status/Overrange
//     PlcTask Inputs/PRG_SL1L0_POWER.fbSL1L0.RTD_South_2.bOverrange <-> RTD Inputs Channel 2/Status/Overrange
//     PlcTask Inputs/PRG_SL1L0_POWER.fbSL1L0.RTD_South_1.bUnderrange <-> RTD Inputs Channel 1/Status/Underrange
//     PlcTask Inputs/PRG_SL1L0_POWER.fbSL1L0.RTD_South_2.bUnderrange <-> RTD Inputs Channel 2/Status/Underrange
//     PlcTask Inputs/PRG_SL1L0_POWER.fbSL1L0.RTD_South_1.iRaw <-> RTD Inputs Channel 1/Value
//     PlcTask Inputs/PRG_SL1L0_POWER.fbSL1L0.RTD_South_2.iRaw <-> RTD Inputs Channel 2/Value
//   lfe_motion Instance <-> PLC Rail (EtherCAT)/Power (EK1200)/PLC Junction 2 (EK1122)/X1 HXR EC1 (EK1100)/EC1 E1 (EK1122)/X1 SL1L0-Power (EK1100)/SL1L0-EL7041-E1
//     PlcTask Inputs/Main.M41.bLimitBackwardEnable <-> STM Status/Status/Digital input 1
//     PlcTask Inputs/Main.M41.bLimitForwardEnable <-> STM Status/Status/Digital input 2
//   lfe_motion Instance <-> PLC Rail (EtherCAT)/Power (EK1200)/PLC Junction 2 (EK1122)/X1 HXR EC1 (EK1100)/EC1 E1 (EK1122)/X1 SL1L0-Power (EK1100)/SL1L0-EL7041-E3
//     PlcTask Inputs/Main.M42.bLimitBackwardEnable <-> STM Status/Status/Digital input 2
//     PlcTask Inputs/Main.M42.bLimitForwardEnable <-> STM Status/Status/Digital input 1
//   lfe_motion Instance <-> PLC Rail (EtherCAT)/Power (EK1200)/PLC Junction 2 (EK1122)/X1 HXR EC1 (EK1100)/EC1 E1 (EK1122)/X1 SL1L0-Power (EK1100)/SL1L0-EL7041-E5
//     PlcTask Inputs/Main.M43.bLimitBackwardEnable <-> STM Status/Status/Digital input 1
//     PlcTask Inputs/Main.M43.bLimitForwardEnable <-> STM Status/Status/Digital input 2
//   lfe_motion Instance <-> PLC Rail (EtherCAT)/Power (EK1200)/PLC Junction 2 (EK1122)/X1 HXR EC1 (EK1100)/EC1 E1 (EK1122)/X1 SL1L0-Power (EK1100)/SL1L0-EL7041-E7
//     PlcTask Inputs/Main.M44.bLimitBackwardEnable <-> STM Status/Status/Digital input 2
//     PlcTask Inputs/Main.M44.bLimitForwardEnable <-> STM Status/Status/Digital input 1
//   lfe_motion Instance <-> PLC Rail (EtherCAT)/Power (EK1200)/PLC Junction 2 (EK1122)/X1 HXR EC1 (EK1100)/EC1 E1 (EK1122)/X2 AT2L0-SOLID (EK1100)/AT2L0-EL7041-01
//     PlcTask Inputs/Main.M1.bLimitBackwardEnable <-> STM Status/Status/Digital input 1
//     PlcTask Inputs/Main.M1.bLimitForwardEnable <-> STM Status/Status/Digital input 2
//     PlcTask Inputs/PRG_AT2L0_SOLID.nM1CoilARaw <-> STM Synchron info data/Info data 1
//     PlcTask Inputs/PRG_AT2L0_SOLID.nM1CoilBRaw <-> STM Synchron info data/Info data 2
//   lfe_motion Instance <-> PLC Rail (EtherCAT)/Power (EK1200)/PLC Junction 2 (EK1122)/X1 HXR EC1 (EK1100)/EC1 E1 (EK1122)/X2 AT2L0-SOLID (EK1100)/AT2L0-EL7041-02
//     PlcTask Inputs/Main.M2.bLimitBackwardEnable <-> STM Status/Status/Digital input 1
//     PlcTask Inputs/Main.M2.bLimitForwardEnable <-> STM Status/Status/Digital input 2
//     PlcTask Inputs/PRG_AT2L0_SOLID.nM2CoilARaw <-> STM Synchron info data/Info data 1
//     PlcTask Inputs/PRG_AT2L0_SOLID.nM2CoilBRaw <-> STM Synchron info data/Info data 2
//   lfe_motion Instance <-> PLC Rail (EtherCAT)/Power (EK1200)/PLC Junction 2 (EK1122)/X1 HXR EC1 (EK1100)/EC1 E1 (EK1122)/X2 AT2L0-SOLID (EK1100)/AT2L0-EL7041-03
//     PlcTask Inputs/Main.M3.bLimitBackwardEnable <-> STM Status/Status/Digital input 1
//     PlcTask Inputs/Main.M3.bLimitForwardEnable <-> STM Status/Status/Digital input 2
//     PlcTask Inputs/PRG_AT2L0_SOLID.nM3CoilARaw <-> STM Synchron info data/Info data 1
//     PlcTask Inputs/PRG_AT2L0_SOLID.nM3CoilBRaw <-> STM Synchron info data/Info data 2
//   lfe_motion Instance <-> PLC Rail (EtherCAT)/Power (EK1200)/PLC Junction 2 (EK1122)/X1 HXR EC1 (EK1100)/EC1 E1 (EK1122)/X2 AT2L0-SOLID (EK1100)/AT2L0-EL7041-04
//     PlcTask Inputs/Main.M4.bLimitBackwardEnable <-> STM Status/Status/Digital input 1
//     PlcTask Inputs/Main.M4.bLimitForwardEnable <-> STM Status/Status/Digital input 2
//     PlcTask Inputs/PRG_AT2L0_SOLID.nM4CoilARaw <-> STM Synchron info data/Info data 1
//     PlcTask Inputs/PRG_AT2L0_SOLID.nM4CoilBRaw <-> STM Synchron info data/Info data 2
//   lfe_motion Instance <-> PLC Rail (EtherCAT)/Power (EK1200)/PLC Junction 2 (EK1122)/X1 HXR EC1 (EK1100)/EC1 E1 (EK1122)/X2 AT2L0-SOLID (EK1100)/AT2L0-EL7041-05
//     PlcTask Inputs/Main.M5.bLimitBackwardEnable <-> STM Status/Status/Digital input 1
//     PlcTask Inputs/Main.M5.bLimitForwardEnable <-> STM Status/Status/Digital input 2
//     PlcTask Inputs/PRG_AT2L0_SOLID.nM5CoilARaw <-> STM Synchron info data/Info data 1
//     PlcTask Inputs/PRG_AT2L0_SOLID.nM5CoilBRaw <-> STM Synchron info data/Info data 2
//   lfe_motion Instance <-> PLC Rail (EtherCAT)/Power (EK1200)/PLC Junction 2 (EK1122)/X1 HXR EC1 (EK1100)/EC1 E1 (EK1122)/X2 AT2L0-SOLID (EK1100)/AT2L0-EL7041-06
//     PlcTask Inputs/Main.M6.bLimitBackwardEnable <-> STM Status/Status/Digital input 1
//     PlcTask Inputs/Main.M6.bLimitForwardEnable <-> STM Status/Status/Digital input 2
//     PlcTask Inputs/PRG_AT2L0_SOLID.nM6CoilARaw <-> STM Synchron info data/Info data 1
//     PlcTask Inputs/PRG_AT2L0_SOLID.nM6CoilBRaw <-> STM Synchron info data/Info data 2
//   lfe_motion Instance <-> PLC Rail (EtherCAT)/Power (EK1200)/PLC Junction 2 (EK1122)/X1 HXR EC1 (EK1100)/EC1 E1 (EK1122)/X2 AT2L0-SOLID (EK1100)/AT2L0-EL7041-07
//     PlcTask Inputs/Main.M7.bLimitBackwardEnable <-> STM Status/Status/Digital input 1
//     PlcTask Inputs/Main.M7.bLimitForwardEnable <-> STM Status/Status/Digital input 2
//     PlcTask Inputs/PRG_AT2L0_SOLID.nM7CoilARaw <-> STM Synchron info data/Info data 1
//     PlcTask Inputs/PRG_AT2L0_SOLID.nM7CoilBRaw <-> STM Synchron info data/Info data 2
//   lfe_motion Instance <-> PLC Rail (EtherCAT)/Power (EK1200)/PLC Junction 2 (EK1122)/X1 HXR EC1 (EK1100)/EC1 E1 (EK1122)/X2 AT2L0-SOLID (EK1100)/AT2L0-EL7041-08
//     PlcTask Inputs/Main.M8.bLimitBackwardEnable <-> STM Status/Status/Digital input 1
//     PlcTask Inputs/Main.M8.bLimitForwardEnable <-> STM Status/Status/Digital input 2
//     PlcTask Inputs/PRG_AT2L0_SOLID.nM8CoilARaw <-> STM Synchron info data/Info data 1
//     PlcTask Inputs/PRG_AT2L0_SOLID.nM8CoilBRaw <-> STM Synchron info data/Info data 2
//   lfe_motion Instance <-> PLC Rail (EtherCAT)/Power (EK1200)/PLC Junction 2 (EK1122)/X1 HXR EC1 (EK1100)/EC1 E1 (EK1122)/X2 AT2L0-SOLID (EK1100)/AT2L0-EL7041-09
//     PlcTask Inputs/Main.M9.bLimitBackwardEnable <-> STM Status/Status/Digital input 1
//     PlcTask Inputs/Main.M9.bLimitForwardEnable <-> STM Status/Status/Digital input 2
//     PlcTask Inputs/PRG_AT2L0_SOLID.nM9CoilARaw <-> STM Synchron info data/Info data 1
//     PlcTask Inputs/PRG_AT2L0_SOLID.nM9CoilBRaw <-> STM Synchron info data/Info data 2
//   lfe_motion Instance <-> PLC Rail (EtherCAT)/Power (EK1200)/PLC Junction 2 (EK1122)/X1 HXR EC1 (EK1100)/EC1 E1 (EK1122)/X2 AT2L0-SOLID (EK1100)/AT2L0-EL7041-10
//     PlcTask Inputs/Main.M10.bLimitBackwardEnable <-> STM Status/Status/Digital input 1
//     PlcTask Inputs/Main.M10.bLimitForwardEnable <-> STM Status/Status/Digital input 2
//     PlcTask Inputs/PRG_AT2L0_SOLID.nM10CoilARaw <-> STM Synchron info data/Info data 1
//     PlcTask Inputs/PRG_AT2L0_SOLID.nM10CoilBRaw <-> STM Synchron info data/Info data 2
//   lfe_motion Instance <-> PLC Rail (EtherCAT)/Power (EK1200)/PLC Junction 2 (EK1122)/X1 HXR EC1 (EK1100)/EC1 E1 (EK1122)/X2 AT2L0-SOLID (EK1100)/AT2L0-EL7041-11
//     PlcTask Inputs/Main.M11.bLimitBackwardEnable <-> STM Status/Status/Digital input 1
//     PlcTask Inputs/Main.M11.bLimitForwardEnable <-> STM Status/Status/Digital input 2
//     PlcTask Inputs/PRG_AT2L0_SOLID.nM11CoilARaw <-> STM Synchron info data/Info data 1
//     PlcTask Inputs/PRG_AT2L0_SOLID.nM11CoilBRaw <-> STM Synchron info data/Info data 2
//   lfe_motion Instance <-> PLC Rail (EtherCAT)/Power (EK1200)/PLC Junction 2 (EK1122)/X1 HXR EC1 (EK1100)/EC1 E1 (EK1122)/X2 AT2L0-SOLID (EK1100)/AT2L0-EL7041-12
//     PlcTask Inputs/Main.M12.bLimitBackwardEnable <-> STM Status/Status/Digital input 1
//     PlcTask Inputs/Main.M12.bLimitForwardEnable <-> STM Status/Status/Digital input 2
//     PlcTask Inputs/PRG_AT2L0_SOLID.nM12CoilARaw <-> STM Synchron info data/Info data 1
//     PlcTask Inputs/PRG_AT2L0_SOLID.nM12CoilBRaw <-> STM Synchron info data/Info data 2
//   lfe_motion Instance <-> PLC Rail (EtherCAT)/Power (EK1200)/PLC Junction 2 (EK1122)/X1 HXR EC1 (EK1100)/EC1 E1 (EK1122)/X2 AT2L0-SOLID (EK1100)/AT2L0-EL7041-13
//     PlcTask Inputs/Main.M13.bLimitBackwardEnable <-> STM Status/Status/Digital input 1
//     PlcTask Inputs/Main.M13.bLimitForwardEnable <-> STM Status/Status/Digital input 2
//     PlcTask Inputs/PRG_AT2L0_SOLID.nM13CoilARaw <-> STM Synchron info data/Info data 1
//     PlcTask Inputs/PRG_AT2L0_SOLID.nM13CoilBRaw <-> STM Synchron info data/Info data 2
//   lfe_motion Instance <-> PLC Rail (EtherCAT)/Power (EK1200)/PLC Junction 2 (EK1122)/X1 HXR EC1 (EK1100)/EC1 E1 (EK1122)/X2 AT2L0-SOLID (EK1100)/AT2L0-EL7041-14
//     PlcTask Inputs/Main.M14.bLimitBackwardEnable <-> STM Status/Status/Digital input 1
//     PlcTask Inputs/Main.M14.bLimitForwardEnable <-> STM Status/Status/Digital input 2
//     PlcTask Inputs/PRG_AT2L0_SOLID.nM14CoilARaw <-> STM Synchron info data/Info data 1
//     PlcTask Inputs/PRG_AT2L0_SOLID.nM14CoilBRaw <-> STM Synchron info data/Info data 2
//   lfe_motion Instance <-> PLC Rail (EtherCAT)/Power (EK1200)/PLC Junction 2 (EK1122)/X1 HXR EC1 (EK1100)/EC1 E1 (EK1122)/X2 AT2L0-SOLID (EK1100)/AT2L0-EL7041-15
//     PlcTask Inputs/Main.M15.bLimitBackwardEnable <-> STM Status/Status/Digital input 1
//     PlcTask Inputs/Main.M15.bLimitForwardEnable <-> STM Status/Status/Digital input 2
//     PlcTask Inputs/PRG_AT2L0_SOLID.nM15CoilARaw <-> STM Synchron info data/Info data 1
//     PlcTask Inputs/PRG_AT2L0_SOLID.nM15CoilBRaw <-> STM Synchron info data/Info data 2
//   lfe_motion Instance <-> PLC Rail (EtherCAT)/Power (EK1200)/PLC Junction 2 (EK1122)/X1 HXR EC1 (EK1100)/EC1 E1 (EK1122)/X2 AT2L0-SOLID (EK1100)/AT2L0-EL7041-16
//     PlcTask Inputs/Main.M16.bLimitBackwardEnable <-> STM Status/Status/Digital input 1
//     PlcTask Inputs/Main.M16.bLimitForwardEnable <-> STM Status/Status/Digital input 2
//     PlcTask Inputs/PRG_AT2L0_SOLID.nM16CoilARaw <-> STM Synchron info data/Info data 1
//     PlcTask Inputs/PRG_AT2L0_SOLID.nM16CoilBRaw <-> STM Synchron info data/Info data 2
//   lfe_motion Instance <-> PLC Rail (EtherCAT)/Power (EK1200)/PLC Junction 2 (EK1122)/X1 HXR EC1 (EK1100)/EC1 E1 (EK1122)/X2 AT2L0-SOLID (EK1100)/AT2L0-EL7041-17
//     PlcTask Inputs/Main.M17.bLimitBackwardEnable <-> STM Status/Status/Digital input 1
//     PlcTask Inputs/Main.M17.bLimitForwardEnable <-> STM Status/Status/Digital input 2
//     PlcTask Inputs/PRG_AT2L0_SOLID.nM17CoilARaw <-> STM Synchron info data/Info data 1
//     PlcTask Inputs/PRG_AT2L0_SOLID.nM17CoilBRaw <-> STM Synchron info data/Info data 2
//   lfe_motion Instance <-> PLC Rail (EtherCAT)/Power (EK1200)/PLC Junction 2 (EK1122)/X1 HXR EC1 (EK1100)/EC1 E1 (EK1122)/X2 AT2L0-SOLID (EK1100)/AT2L0-EL7041-18
//     PlcTask Inputs/Main.M18.bLimitBackwardEnable <-> STM Status/Status/Digital input 1
//     PlcTask Inputs/Main.M18.bLimitForwardEnable <-> STM Status/Status/Digital input 2
//     PlcTask Inputs/PRG_AT2L0_SOLID.nM18CoilARaw <-> STM Synchron info data/Info data 1
//     PlcTask Inputs/PRG_AT2L0_SOLID.nM18CoilBRaw <-> STM Synchron info data/Info data 2
//   lfe_motion Instance <-> PLC Rail (EtherCAT)/Power (EK1200)/PLC Junction 2 (EK1122)/X1 HXR EC1 (EK1100)/EC1 E1 (EK1122)/X2 AT2L0-SOLID (EK1100)/AT2L0-EL7041-19
//     PlcTask Inputs/Main.M19.bLimitBackwardEnable <-> STM Status/Status/Digital input 1
//     PlcTask Inputs/Main.M19.bLimitForwardEnable <-> STM Status/Status/Digital input 2
//     PlcTask Inputs/PRG_AT2L0_SOLID.nM19CoilARaw <-> STM Synchron info data/Info data 1
//     PlcTask Inputs/PRG_AT2L0_SOLID.nM19CoilBRaw <-> STM Synchron info data/Info data 2
//   lfe_motion Instance <-> PLC Rail (EtherCAT)/Power (EK1200)/PLC Junction 2 (EK1122)/X1 HXR EC1 (EK1100)/EC1 E2 (EK1122)/X1 IM2L0-XTES (EK1100)/IM2L0-EL1088
//     PlcTask Inputs/Main.M25.bHome <-> Channel 2/Input
//     PlcTask Inputs/Main.M26.bHome <-> Channel 4/Input
//     PlcTask Inputs/PRG_IM2L0_XTES.fbIM2L0.bFocusEndBwd <-> Channel 4/Input
//     PlcTask Inputs/PRG_IM2L0_XTES.fbIM2L0.bFocusEndFwd <-> Channel 3/Input
//     PlcTask Inputs/PRG_IM2L0_XTES.fbIM2L0.bZoomEndBwd <-> Channel 2/Input
//     PlcTask Inputs/PRG_IM2L0_XTES.fbIM2L0.bZoomEndFwd <-> Channel 1/Input
//   lfe_motion Instance <-> PLC Rail (EtherCAT)/Power (EK1200)/PLC Junction 2 (EK1122)/X1 HXR EC1 (EK1100)/EC1 E2 (EK1122)/X1 IM2L0-XTES (EK1100)/IM2L0-EL2004
//     PlcTask Outputs/Main.M24.bBrakeRelease <-> Channel 1/Output
//     PlcTask Outputs/PRG_IM2L0_XTES.fbIM2L0.fbLED.bLEDPower <-> Channel 3/Output
//     PlcTask Outputs/PRG_IM2L0_XTES.fbIM2L0.fbOpal.bOpalPower <-> Channel 2/Output
//   lfe_motion Instance <-> PLC Rail (EtherCAT)/Power (EK1200)/PLC Junction 2 (EK1122)/X1 HXR EC1 (EK1100)/EC1 E2 (EK1122)/X1 IM2L0-XTES (EK1100)/IM2L0-EL6002
//     PlcTask Inputs/PRG_IM2L0_XTES.stEL6In/D[{0..21}] <-> COM TxPDO-Map Inputs Channel 1/Data In {0..21}  (22 links)
//     PlcTask Inputs/PRG_IM2L0_XTES.stEL6In/Status <-> COM TxPDO-Map Inputs Channel 1/Status
//     PlcTask Outputs/PRG_IM2L0_XTES.stEL6Out/Ctrl <-> COM RxPDO-Map Outputs Channel 1/Ctrl
//     PlcTask Outputs/PRG_IM2L0_XTES.stEL6Out/D[{0..21}] <-> COM RxPDO-Map Outputs Channel 1/Data Out {0..21}  (22 links)
//   lfe_motion Instance <-> PLC Rail (EtherCAT)/Power (EK1200)/PLC Junction 2 (EK1122)/X1 HXR EC1 (EK1100)/EC1 E2 (EK1122)/X1 IM2L0-XTES (EK1100)/IM2L0-EL7041
//     PlcTask Inputs/PRG_IM2L0_XTES.bDefectiveLimitSwitch <-> STM Status/Status/Digital input 1
//   lfe_motion Instance <-> PLC Rail (EtherCAT)/Power (EK1200)/PLC Junction 2 (EK1122)/X1 HXR EC1 (EK1100)/EC1 E2 (EK1122)/X2 SL2L0-Power (EK1100)/SL2L0-EL3202-E10
//     PlcTask Inputs/PRG_SL2L0_POWER.fbSL2L0.RTD_North_1.bError <-> RTD Inputs Channel 1/Status/Error
//     PlcTask Inputs/PRG_SL2L0_POWER.fbSL2L0.RTD_North_1.iRaw <-> RTD Inputs Channel 1/Value
//     PlcTask Inputs/PRG_SL2L0_POWER.fbSL2L0.RTD_TOP_1.bError <-> RTD Inputs Channel 1/Status/Error
//     PlcTask Inputs/PRG_SL2L0_POWER.fbSL2L0.RTD_TOP_2.bError <-> RTD Inputs Channel 2/Status/Error
//     PlcTask Inputs/PRG_SL2L0_POWER.fbSL2L0.RTD_TOP_1.bOverrange <-> RTD Inputs Channel 1/Status/Overrange
//     PlcTask Inputs/PRG_SL2L0_POWER.fbSL2L0.RTD_TOP_2.bOverrange <-> RTD Inputs Channel 2/Status/Overrange
//     PlcTask Inputs/PRG_SL2L0_POWER.fbSL2L0.RTD_TOP_1.bUnderrange <-> RTD Inputs Channel 1/Status/Underrange
//     PlcTask Inputs/PRG_SL2L0_POWER.fbSL2L0.RTD_TOP_2.bUnderrange <-> RTD Inputs Channel 2/Status/Underrange
//     PlcTask Inputs/PRG_SL2L0_POWER.fbSL2L0.RTD_TOP_1.iRaw <-> RTD Inputs Channel 1/Value
//     PlcTask Inputs/PRG_SL2L0_POWER.fbSL2L0.RTD_TOP_2.iRaw <-> RTD Inputs Channel 2/Value
//   lfe_motion Instance <-> PLC Rail (EtherCAT)/Power (EK1200)/PLC Junction 2 (EK1122)/X1 HXR EC1 (EK1100)/EC1 E2 (EK1122)/X2 SL2L0-Power (EK1100)/SL2L0-EL3202-E11
//     PlcTask Inputs/PRG_SL2L0_POWER.fbSL2L0.RTD_North_1.bOverrange <-> RTD Inputs Channel 1/Status/Overrange
//     PlcTask Inputs/PRG_SL2L0_POWER.fbSL2L0.RTD_North_2.bOverrange <-> RTD Inputs Channel 2/Status/Overrange
//     PlcTask Inputs/PRG_SL2L0_POWER.fbSL2L0.RTD_North_1.bUnderrange <-> RTD Inputs Channel 1/Status/Underrange
//     PlcTask Inputs/PRG_SL2L0_POWER.fbSL2L0.RTD_North_2.bUnderrange <-> RTD Inputs Channel 2/Status/Underrange
//     PlcTask Inputs/PRG_SL2L0_POWER.fbSL2L0.RTD_North_2.bError <-> RTD Inputs Channel 2/Status/Error
//     PlcTask Inputs/PRG_SL2L0_POWER.fbSL2L0.RTD_North_2.iRaw <-> RTD Inputs Channel 2/Value
//   lfe_motion Instance <-> PLC Rail (EtherCAT)/Power (EK1200)/PLC Junction 2 (EK1122)/X1 HXR EC1 (EK1100)/EC1 E2 (EK1122)/X2 SL2L0-Power (EK1100)/SL2L0-EL3202-E8
//     PlcTask Inputs/PRG_SL2L0_POWER.fbSL2L0.RTD_Bottom_1.bError <-> RTD Inputs Channel 1/Status/Error
//     PlcTask Inputs/PRG_SL2L0_POWER.fbSL2L0.RTD_Bottom_2.bError <-> RTD Inputs Channel 2/Status/Error
//     PlcTask Inputs/PRG_SL2L0_POWER.fbSL2L0.RTD_Bottom_1.bOverrange <-> RTD Inputs Channel 1/Status/Overrange
//     PlcTask Inputs/PRG_SL2L0_POWER.fbSL2L0.RTD_Bottom_2.bOverrange <-> RTD Inputs Channel 2/Status/Overrange
//     PlcTask Inputs/PRG_SL2L0_POWER.fbSL2L0.RTD_Bottom_1.bUnderrange <-> RTD Inputs Channel 1/Status/Underrange
//     PlcTask Inputs/PRG_SL2L0_POWER.fbSL2L0.RTD_Bottom_2.bUnderrange <-> RTD Inputs Channel 2/Status/Underrange
//     PlcTask Inputs/PRG_SL2L0_POWER.fbSL2L0.RTD_Bottom_1.iRaw <-> RTD Inputs Channel 1/Value
//     PlcTask Inputs/PRG_SL2L0_POWER.fbSL2L0.RTD_Bottom_2.iRaw <-> RTD Inputs Channel 2/Value
//   lfe_motion Instance <-> PLC Rail (EtherCAT)/Power (EK1200)/PLC Junction 2 (EK1122)/X1 HXR EC1 (EK1100)/EC1 E2 (EK1122)/X2 SL2L0-Power (EK1100)/SL2L0-EL3202-E9
//     PlcTask Inputs/PRG_SL2L0_POWER.fbSL2L0.RTD_South_1.bError <-> RTD Inputs Channel 1/Status/Error
//     PlcTask Inputs/PRG_SL2L0_POWER.fbSL2L0.RTD_South_2.bError <-> RTD Inputs Channel 2/Status/Error
//     PlcTask Inputs/PRG_SL2L0_POWER.fbSL2L0.RTD_South_1.bOverrange <-> RTD Inputs Channel 1/Status/Overrange
//     PlcTask Inputs/PRG_SL2L0_POWER.fbSL2L0.RTD_South_2.bOverrange <-> RTD Inputs Channel 2/Status/Overrange
//     PlcTask Inputs/PRG_SL2L0_POWER.fbSL2L0.RTD_South_1.bUnderrange <-> RTD Inputs Channel 1/Status/Underrange
//     PlcTask Inputs/PRG_SL2L0_POWER.fbSL2L0.RTD_South_2.bUnderrange <-> RTD Inputs Channel 2/Status/Underrange
//     PlcTask Inputs/PRG_SL2L0_POWER.fbSL2L0.RTD_South_1.iRaw <-> RTD Inputs Channel 1/Value
//     PlcTask Inputs/PRG_SL2L0_POWER.fbSL2L0.RTD_South_2.iRaw <-> RTD Inputs Channel 2/Value
//   lfe_motion Instance <-> PLC Rail (EtherCAT)/Power (EK1200)/PLC Junction 2 (EK1122)/X1 HXR EC1 (EK1100)/EC1 E2 (EK1122)/X2 SL2L0-Power (EK1100)/SL2L0-EL7041-E1
//     PlcTask Inputs/Main.M45.bLimitBackwardEnable <-> STM Status/Status/Digital input 1
//     PlcTask Inputs/Main.M45.bLimitForwardEnable <-> STM Status/Status/Digital input 2
//   lfe_motion Instance <-> PLC Rail (EtherCAT)/Power (EK1200)/PLC Junction 2 (EK1122)/X1 HXR EC1 (EK1100)/EC1 E2 (EK1122)/X2 SL2L0-Power (EK1100)/SL2L0-EL7041-E3
//     PlcTask Inputs/Main.M46.bLimitBackwardEnable <-> STM Status/Status/Digital input 2
//     PlcTask Inputs/Main.M46.bLimitForwardEnable <-> STM Status/Status/Digital input 1
//   lfe_motion Instance <-> PLC Rail (EtherCAT)/Power (EK1200)/PLC Junction 2 (EK1122)/X1 HXR EC1 (EK1100)/EC1 E2 (EK1122)/X2 SL2L0-Power (EK1100)/SL2L0-EL7041-E5
//     PlcTask Inputs/Main.M47.bLimitBackwardEnable <-> STM Status/Status/Digital input 1
//     PlcTask Inputs/Main.M47.bLimitForwardEnable <-> STM Status/Status/Digital input 2
//   lfe_motion Instance <-> PLC Rail (EtherCAT)/Power (EK1200)/PLC Junction 2 (EK1122)/X1 HXR EC1 (EK1100)/EC1 E2 (EK1122)/X2 SL2L0-Power (EK1100)/SL2L0-EL7041-E7
//     PlcTask Inputs/Main.M48.bLimitBackwardEnable <-> STM Status/Status/Digital input 2
//     PlcTask Inputs/Main.M48.bLimitForwardEnable <-> STM Status/Status/Digital input 1
//   lfe_motion Instance <-> PLC Rail (EtherCAT)/Power (EK1200)/PLC Junction 2 (EK1122)/X1 HXR EC1 (EK1100)/EC1 E3 (EK1122)/X1 PF1L0-WFS (EK1100)/PF1L0-EL2004
//     PlcTask Outputs/Main.M31.bBrakeRelease <-> Channel 1/Output
//   lfe_motion Instance <-> PLC Rail (EtherCAT)/Power (EK1200)/PLC Junction 2 (EK1122)/X1 HXR EC1 (EK1100)/EC1 E3 (EK1122)/X1 PF1L0-WFS (EK1100)/PF1L0-EL3314
//     PlcTask Inputs/PRG_PF1L0_WFS.fbPF1L0.fbThermoCouple1.bError <-> TC Inputs Channel 1/Status/Error
//     PlcTask Inputs/PRG_PF1L0_WFS.fbPF1L0.fbThermoCouple2.bError <-> TC Inputs Channel 2/Status/Error
//     PlcTask Inputs/PRG_PF1L0_WFS.fbPF1L0.fbThermoCouple1.bOverrange <-> TC Inputs Channel 1/Status/Overrange
//     PlcTask Inputs/PRG_PF1L0_WFS.fbPF1L0.fbThermoCouple2.bOverrange <-> TC Inputs Channel 2/Status/Overrange
//     PlcTask Inputs/PRG_PF1L0_WFS.fbPF1L0.fbThermoCouple1.bUnderrange <-> TC Inputs Channel 1/Status/Underrange
//     PlcTask Inputs/PRG_PF1L0_WFS.fbPF1L0.fbThermoCouple2.bUnderrange <-> TC Inputs Channel 2/Status/Underrange
//     PlcTask Inputs/PRG_PF1L0_WFS.fbPF1L0.fbThermoCouple1.iRaw <-> TC Inputs Channel 1/Value
//     PlcTask Inputs/PRG_PF1L0_WFS.fbPF1L0.fbThermoCouple2.iRaw <-> TC Inputs Channel 2/Value
//   lfe_motion Instance <-> PLC Rail (EtherCAT)/Power (EK1200)/PLC Junction 2 (EK1122)/X1 HXR EC1 (EK1100)/EC1 E3 (EK1122)/X1 PF1L0-WFS (EK1100)/PF1L0-EL5042
//     PlcTask Inputs/Main.M31.nRawEncoderULINT <-> FB Inputs Channel 2/Position
//     PlcTask Inputs/Main.M32.nRawEncoderULINT <-> FB Inputs Channel 1/Position
//   lfe_motion Instance <-> PLC Rail (EtherCAT)/Power (EK1200)/PLC Junction 2 (EK1122)/X1 HXR EC1 (EK1100)/EC1 E3 (EK1122)/X1 PF1L0-WFS (EK1100)/PF1L0-EL7041-01
//     PlcTask Inputs/Main.M31.bLimitBackwardEnable <-> STM Status/Status/Digital input 2
//     PlcTask Inputs/Main.M31.bLimitForwardEnable <-> STM Status/Status/Digital input 1
//   lfe_motion Instance <-> PLC Rail (EtherCAT)/Power (EK1200)/PLC Junction 2 (EK1122)/X1 HXR EC1 (EK1100)/EC1 E3 (EK1122)/X2_0 SP1L0-KMONO_MOTOR (EK1100)/SP1L0-EL7041-E2-MOTORS
//     PlcTask Inputs/Main.M50.bLimitBackwardEnable <-> STM Status/Status/Digital input 1
//     PlcTask Inputs/Main.M50.bLimitForwardEnable <-> STM Status/Status/Digital input 2
//   lfe_motion Instance <-> PLC Rail (EtherCAT)/Power (EK1200)/PLC Junction 2 (EK1122)/X1 HXR EC1 (EK1100)/EC1 E3 (EK1122)/X2_0 SP1L0-KMONO_MOTOR (EK1100)/SP1L0-EL7041-E3-MOTORS
//     PlcTask Inputs/Main.M51.bLimitBackwardEnable <-> STM Status/Status/Digital input 1
//     PlcTask Inputs/Main.M51.bLimitForwardEnable <-> STM Status/Status/Digital input 2
//   lfe_motion Instance <-> PLC Rail (EtherCAT)/Power (EK1200)/PLC Junction 2 (EK1122)/X1 HXR EC1 (EK1100)/EC1 E3 (EK1122)/X2_0 SP1L0-KMONO_MOTOR (EK1100)/SP1L0-EL7041-E4-MOTORS
//     PlcTask Inputs/Main.M52.bLimitBackwardEnable <-> STM Status/Status/Digital input 2
//     PlcTask Inputs/Main.M52.bLimitForwardEnable <-> STM Status/Status/Digital input 1
//   lfe_motion Instance <-> PLC Rail (EtherCAT)/Power (EK1200)/PLC Junction 2 (EK1122)/X1 HXR EC1 (EK1100)/EC1 E3 (EK1122)/X2_0 SP1L0-KMONO_MOTOR (EK1100)/SP1L0-EL7041-E5-MOTORS
//     PlcTask Inputs/Main.M53.bLimitBackwardEnable <-> STM Status/Status/Digital input 1
//     PlcTask Inputs/Main.M53.bLimitForwardEnable <-> STM Status/Status/Digital input 2
//   lfe_motion Instance <-> PLC Rail (EtherCAT)/Power (EK1200)/PLC Junction 2 (EK1122)/X1 HXR EC1 (EK1100)/EC1 E3 (EK1122)/X2_0 SP1L0-KMONO_MOTOR (EK1100)/SP1L0-EL7041-E6-MOTORS
//     PlcTask Inputs/Main.M54.bLimitBackwardEnable <-> STM Status/Status/Digital input 2
//     PlcTask Inputs/Main.M54.bLimitForwardEnable <-> STM Status/Status/Digital input 1
//   lfe_motion Instance <-> PLC Rail (EtherCAT)/Power (EK1200)/PLC Junction 2 (EK1122)/X2 HXR EC2 (EK1100)/EC2 E1 (EK1122)/X1 IM3L0-PPM (EK1100)/IM3L0-EL2004
//     PlcTask Outputs/Main.M27.bBrakeRelease <-> Channel 1/Output
//     PlcTask Outputs/PRG_IM3L0_PPM.fbIM3L0.fbGige.bGigePower <-> Channel 2/Output
//   lfe_motion Instance <-> PLC Rail (EtherCAT)/Power (EK1200)/PLC Junction 2 (EK1122)/X2 HXR EC2 (EK1100)/EC2 E1 (EK1122)/X1 IM3L0-PPM (EK1100)/IM3L0-EL3062
//     PlcTask Inputs/PRG_IM3L0_PPM.fbIM3L0.fbPowerMeter.iVoltageINT <-> AI Standard Channel 1/Value
//   lfe_motion Instance <-> PLC Rail (EtherCAT)/Power (EK1200)/PLC Junction 2 (EK1122)/X2 HXR EC2 (EK1100)/EC2 E1 (EK1122)/X1 IM3L0-PPM (EK1100)/IM3L0-EL3314
//     PlcTask Inputs/PRG_IM3L0_PPM.fbIM3L0.fbPowerMeter.fbThermoCouple.bError <-> TC Inputs Channel 1/Status/Error
//     PlcTask Inputs/PRG_IM3L0_PPM.fbIM3L0.fbPowerMeter.fbThermoCouple.bOverrange <-> TC Inputs Channel 1/Status/Overrange
//     PlcTask Inputs/PRG_IM3L0_PPM.fbIM3L0.fbPowerMeter.fbThermoCouple.bUnderrange <-> TC Inputs Channel 1/Status/Underrange
//     PlcTask Inputs/PRG_IM3L0_PPM.fbIM3L0.fbPowerMeter.fbThermoCouple.iRaw <-> TC Inputs Channel 1/Value
//     PlcTask Inputs/PRG_IM3L0_PPM.fbIM3L0.fbYagThermoCouple.bError <-> TC Inputs Channel 2/Status/Error
//     PlcTask Inputs/PRG_IM3L0_PPM.fbIM3L0.fbYagThermoCouple.bOverrange <-> TC Inputs Channel 2/Status/Overrange
//     PlcTask Inputs/PRG_IM3L0_PPM.fbIM3L0.fbYagThermoCouple.bUnderrange <-> TC Inputs Channel 2/Status/Underrange
//     PlcTask Inputs/PRG_IM3L0_PPM.fbIM3L0.fbYagThermoCouple.iRaw <-> TC Inputs Channel 2/Value
//   lfe_motion Instance <-> PLC Rail (EtherCAT)/Power (EK1200)/PLC Junction 2 (EK1122)/X2 HXR EC2 (EK1100)/EC2 E1 (EK1122)/X1 IM3L0-PPM (EK1100)/IM3L0-EL4004
//     PlcTask Outputs/PRG_IM3L0_PPM.fbIM3L0.fbGige.iIlluminatorINT <-> AO Outputs Channel 1/Analog output
//   lfe_motion Instance <-> PLC Rail (EtherCAT)/Power (EK1200)/PLC Junction 2 (EK1122)/X2 HXR EC2 (EK1100)/EC2 E1 (EK1122)/X1 IM3L0-PPM (EK1100)/IM3L0-EL7041
//     PlcTask Inputs/Main.M27.bLimitBackwardEnable <-> STM Status/Status/Digital input 2
//     PlcTask Inputs/Main.M27.bLimitForwardEnable <-> STM Status/Status/Digital input 1
//   lfe_motion Instance <-> PLC Rail (EtherCAT)/Power (EK1200)/PLC Junction 2 (EK1122)/X2 HXR EC2 (EK1100)/EC2 E1 (EK1122)/X2 IM1L1-PPM (EK1100)/IM1L1-EL2004
//     PlcTask Outputs/Main.M23.bBrakeRelease <-> Channel 1/Output
//     PlcTask Outputs/PRG_IM1L1_PPM.fbIM1L1.fbGige.bGigePower <-> Channel 2/Output
//   lfe_motion Instance <-> PLC Rail (EtherCAT)/Power (EK1200)/PLC Junction 2 (EK1122)/X2 HXR EC2 (EK1100)/EC2 E1 (EK1122)/X2 IM1L1-PPM (EK1100)/IM1L1-EL3062
//     PlcTask Inputs/PRG_IM1L1_PPM.fbIM1L1.fbPowerMeter.iVoltageINT <-> AI Standard Channel 1/Value
//   lfe_motion Instance <-> PLC Rail (EtherCAT)/Power (EK1200)/PLC Junction 2 (EK1122)/X2 HXR EC2 (EK1100)/EC2 E1 (EK1122)/X2 IM1L1-PPM (EK1100)/IM1L1-EL3314
//     PlcTask Inputs/PRG_IM1L1_PPM.fbIM1L1.fbPowerMeter.fbThermoCouple.bError <-> TC Inputs Channel 1/Status/Error
//     PlcTask Inputs/PRG_IM1L1_PPM.fbIM1L1.fbPowerMeter.fbThermoCouple.bOverrange <-> TC Inputs Channel 1/Status/Overrange
//     PlcTask Inputs/PRG_IM1L1_PPM.fbIM1L1.fbPowerMeter.fbThermoCouple.bUnderrange <-> TC Inputs Channel 1/Status/Underrange
//     PlcTask Inputs/PRG_IM1L1_PPM.fbIM1L1.fbPowerMeter.fbThermoCouple.iRaw <-> TC Inputs Channel 1/Value
//     PlcTask Inputs/PRG_IM1L1_PPM.fbIM1L1.fbYagThermoCouple.bError <-> TC Inputs Channel 2/Status/Error
//     PlcTask Inputs/PRG_IM1L1_PPM.fbIM1L1.fbYagThermoCouple.bOverrange <-> TC Inputs Channel 2/Status/Overrange
//     PlcTask Inputs/PRG_IM1L1_PPM.fbIM1L1.fbYagThermoCouple.bUnderrange <-> TC Inputs Channel 2/Status/Underrange
//     PlcTask Inputs/PRG_IM1L1_PPM.fbIM1L1.fbYagThermoCouple.iRaw <-> TC Inputs Channel 2/Value
//   lfe_motion Instance <-> PLC Rail (EtherCAT)/Power (EK1200)/PLC Junction 2 (EK1122)/X2 HXR EC2 (EK1100)/EC2 E1 (EK1122)/X2 IM1L1-PPM (EK1100)/IM1L1-EL4004
//     PlcTask Outputs/PRG_IM1L1_PPM.fbIM1L1.fbGige.iIlluminatorINT <-> AO Outputs Channel 1/Analog output
//   lfe_motion Instance <-> PLC Rail (EtherCAT)/Power (EK1200)/PLC Junction 2 (EK1122)/X2 HXR EC2 (EK1100)/EC2 E1 (EK1122)/X2 IM1L1-PPM (EK1100)/IM1L1-EL7041
//     PlcTask Inputs/Main.M23.bLimitBackwardEnable <-> STM Status/Status/Digital input 2
//     PlcTask Inputs/Main.M23.bLimitForwardEnable <-> STM Status/Status/Digital input 1
//   lfe_motion Instance <-> PLC Rail (EtherCAT)/Power (EK1200)/PLC Junction 2 (EK1122)/X2 HXR EC2 (EK1100)/EC2 E2 (EK1122)/X1 IM4L0-XTES (EK1100)/IM4L0-EL1088
//     PlcTask Inputs/Main.M29.bHome <-> Channel 2/Input
//     PlcTask Inputs/Main.M30.bHome <-> Channel 4/Input
//     PlcTask Inputs/PRG_IM4L0_XTES.fbIM4L0.bFocusEndBwd <-> Channel 4/Input
//     PlcTask Inputs/PRG_IM4L0_XTES.fbIM4L0.bFocusEndFwd <-> Channel 3/Input
//     PlcTask Inputs/PRG_IM4L0_XTES.fbIM4L0.bZoomEndBwd <-> Channel 2/Input
//     PlcTask Inputs/PRG_IM4L0_XTES.fbIM4L0.bZoomEndFwd <-> Channel 1/Input
//   lfe_motion Instance <-> PLC Rail (EtherCAT)/Power (EK1200)/PLC Junction 2 (EK1122)/X2 HXR EC2 (EK1100)/EC2 E2 (EK1122)/X1 IM4L0-XTES (EK1100)/IM4L0-EL2004
//     PlcTask Outputs/Main.M28.bBrakeRelease <-> Channel 1/Output
//     PlcTask Outputs/PRG_IM4L0_XTES.bIM4L0_SCRP_LED_01 <-> Channel 4/Output
//     PlcTask Outputs/PRG_IM4L0_XTES.fbIM4L0.fbLED.bLEDPower <-> Channel 3/Output
//     PlcTask Outputs/PRG_IM4L0_XTES.fbIM4L0.fbOpal.bOpalPower <-> Channel 2/Output
//   lfe_motion Instance <-> PLC Rail (EtherCAT)/Power (EK1200)/PLC Junction 2 (EK1122)/X2 HXR EC2 (EK1100)/EC2 E2 (EK1122)/X1 IM4L0-XTES (EK1100)/IM4L0-EL6002
//     PlcTask Inputs/PRG_IM4L0_XTES.stEL6In/D[{0..21}] <-> COM TxPDO-Map Inputs Channel 1/Data In {0..21}  (22 links)
//     PlcTask Inputs/PRG_IM4L0_XTES.stEL6In/Status <-> COM TxPDO-Map Inputs Channel 1/Status
//     PlcTask Outputs/PRG_IM4L0_XTES.stEL6Out/Ctrl <-> COM RxPDO-Map Outputs Channel 1/Ctrl
//     PlcTask Outputs/PRG_IM4L0_XTES.stEL6Out/D[{0..21}] <-> COM RxPDO-Map Outputs Channel 1/Data Out {0..21}  (22 links)
//   lfe_motion Instance <-> PLC Rail (EtherCAT)/Power (EK1200)/PLC Junction 2 (EK1122)/X2 HXR EC2 (EK1100)/EC2 E2 (EK1122)/X1 IM4L0-XTES (EK1100)/IM4L0-EL7041
//     PlcTask Inputs/Main.M28.bLimitForwardEnable <-> STM Status/Status/Digital input 1
//   lfe_motion Instance <-> PLC Rail (EtherCAT)/Power (EK1200)/PMPS_FFO
//     PlcTask Outputs/GVL.fbFastFaultOutput1.q_xFastFaultOut <-> Channel 1/Output
//     PlcTask Outputs/GVL.fbFastFaultOutput2.q_xFastFaultOut <-> Channel 2/Output
//   lfe_motion Instance <-> PLC Rail (EtherCAT)/Power (EK1200)/PMPS_PRE
//     PlcTask Inputs/GVL.rReqTrans <-> IO Inputs/SattArrayReq
//     PlcTask Inputs/PRG_3_PMPS_POST.fbArbiterIO.i_stCurrentBP <-> IO Inputs/CurrentBP
//     PlcTask Inputs/PRG_3_PMPS_POST.fbArbiterIO.xTxPDO_state <-> SYNC Inputs/TxPDO state
//     PlcTask Inputs/PRG_3_PMPS_POST.fbArbiterIO.xTxPDO_toggle <-> SYNC Inputs/TxPDO toggle
//     PlcTask Outputs/GVL.rCurTrans <-> IO Outputs/SattArrayStatus
//     PlcTask Outputs/PRG_3_PMPS_POST.fbArbiterIO.q_stRequestedBP <-> IO Outputs/RequestedBP
//   lfe_motion Instance <-> NC-Task 1 SAF/Axes/Axis 1
//     PlcTask Inputs/Main.M1.Axis.NcToPlc <-> Outputs/ToPlc
//     PlcTask Outputs/Main.M1.Axis.PlcToNc <-> Inputs/FromPlc
//   lfe_motion Instance <-> NC-Task 1 SAF/Axes/Axis 10
//     PlcTask Inputs/Main.M10.Axis.NcToPlc <-> Outputs/ToPlc
//     PlcTask Outputs/Main.M10.Axis.PlcToNc <-> Inputs/FromPlc
//   lfe_motion Instance <-> NC-Task 1 SAF/Axes/Axis 11
//     PlcTask Inputs/Main.M11.Axis.NcToPlc <-> Outputs/ToPlc
//     PlcTask Outputs/Main.M11.Axis.PlcToNc <-> Inputs/FromPlc
//   lfe_motion Instance <-> NC-Task 1 SAF/Axes/Axis 12
//     PlcTask Inputs/Main.M12.Axis.NcToPlc <-> Outputs/ToPlc
//     PlcTask Outputs/Main.M12.Axis.PlcToNc <-> Inputs/FromPlc
//   lfe_motion Instance <-> NC-Task 1 SAF/Axes/Axis 13
//     PlcTask Inputs/Main.M13.Axis.NcToPlc <-> Outputs/ToPlc
//     PlcTask Outputs/Main.M13.Axis.PlcToNc <-> Inputs/FromPlc
//   lfe_motion Instance <-> NC-Task 1 SAF/Axes/Axis 14
//     PlcTask Inputs/Main.M14.Axis.NcToPlc <-> Outputs/ToPlc
//     PlcTask Outputs/Main.M14.Axis.PlcToNc <-> Inputs/FromPlc
//   lfe_motion Instance <-> NC-Task 1 SAF/Axes/Axis 15
//     PlcTask Inputs/Main.M15.Axis.NcToPlc <-> Outputs/ToPlc
//     PlcTask Outputs/Main.M15.Axis.PlcToNc <-> Inputs/FromPlc
//   lfe_motion Instance <-> NC-Task 1 SAF/Axes/Axis 16
//     PlcTask Inputs/Main.M16.Axis.NcToPlc <-> Outputs/ToPlc
//     PlcTask Outputs/Main.M16.Axis.PlcToNc <-> Inputs/FromPlc
//   lfe_motion Instance <-> NC-Task 1 SAF/Axes/Axis 17
//     PlcTask Inputs/Main.M17.Axis.NcToPlc <-> Outputs/ToPlc
//     PlcTask Outputs/Main.M17.Axis.PlcToNc <-> Inputs/FromPlc
//   lfe_motion Instance <-> NC-Task 1 SAF/Axes/Axis 18
//     PlcTask Inputs/Main.M18.Axis.NcToPlc <-> Outputs/ToPlc
//     PlcTask Outputs/Main.M18.Axis.PlcToNc <-> Inputs/FromPlc
//   lfe_motion Instance <-> NC-Task 1 SAF/Axes/Axis 19
//     PlcTask Inputs/Main.M19.Axis.NcToPlc <-> Outputs/ToPlc
//     PlcTask Outputs/Main.M19.Axis.PlcToNc <-> Inputs/FromPlc
//   lfe_motion Instance <-> NC-Task 1 SAF/Axes/Axis 2
//     PlcTask Inputs/Main.M2.Axis.NcToPlc <-> Outputs/ToPlc
//     PlcTask Outputs/Main.M2.Axis.PlcToNc <-> Inputs/FromPlc
//   lfe_motion Instance <-> NC-Task 1 SAF/Axes/Axis 20 IM1L0-XTES-MMS
//     PlcTask Inputs/Main.M20.Axis.NcToPlc <-> Outputs/ToPlc
//     PlcTask Outputs/Main.M20.Axis.PlcToNc <-> Inputs/FromPlc
//   lfe_motion Instance <-> NC-Task 1 SAF/Axes/Axis 21 IM1L0-XTES-CLZ
//     PlcTask Inputs/Main.M21.Axis.NcToPlc <-> Outputs/ToPlc
//     PlcTask Outputs/Main.M21.Axis.PlcToNc <-> Inputs/FromPlc
//   lfe_motion Instance <-> NC-Task 1 SAF/Axes/Axis 22 IM1L0-XTES-CLF
//     PlcTask Inputs/Main.M22.Axis.NcToPlc <-> Outputs/ToPlc
//     PlcTask Outputs/Main.M22.Axis.PlcToNc <-> Inputs/FromPlc
//   lfe_motion Instance <-> NC-Task 1 SAF/Axes/Axis 23 IM1L1-PPM-MMS
//     PlcTask Inputs/Main.M23.Axis.NcToPlc <-> Outputs/ToPlc
//     PlcTask Outputs/Main.M23.Axis.PlcToNc <-> Inputs/FromPlc
//   lfe_motion Instance <-> NC-Task 1 SAF/Axes/Axis 24 IM2L0-XTES-MMS
//     PlcTask Inputs/Main.M24.Axis.NcToPlc <-> Outputs/ToPlc
//     PlcTask Outputs/Main.M24.Axis.PlcToNc <-> Inputs/FromPlc
//   lfe_motion Instance <-> NC-Task 1 SAF/Axes/Axis 25 IM2L0-XTES-CLZ
//     PlcTask Inputs/Main.M25.Axis.NcToPlc <-> Outputs/ToPlc
//     PlcTask Outputs/Main.M25.Axis.PlcToNc <-> Inputs/FromPlc
//   lfe_motion Instance <-> NC-Task 1 SAF/Axes/Axis 26 IM2L0-XTES-CLF
//     PlcTask Inputs/Main.M26.Axis.NcToPlc <-> Outputs/ToPlc
//     PlcTask Outputs/Main.M26.Axis.PlcToNc <-> Inputs/FromPlc
//   lfe_motion Instance <-> NC-Task 1 SAF/Axes/Axis 27 IM3L0-PPM-MMS
//     PlcTask Inputs/Main.M27.Axis.NcToPlc <-> Outputs/ToPlc
//     PlcTask Outputs/Main.M27.Axis.PlcToNc <-> Inputs/FromPlc
//   lfe_motion Instance <-> NC-Task 1 SAF/Axes/Axis 28 IM4L0-XTES-MMS
//     PlcTask Inputs/Main.M28.Axis.NcToPlc <-> Outputs/ToPlc
//     PlcTask Outputs/Main.M28.Axis.PlcToNc <-> Inputs/FromPlc
//   lfe_motion Instance <-> NC-Task 1 SAF/Axes/Axis 29 IM4L0-XTES-CLZ
//     PlcTask Inputs/Main.M29.Axis.NcToPlc <-> Outputs/ToPlc
//     PlcTask Outputs/Main.M29.Axis.PlcToNc <-> Inputs/FromPlc
//   lfe_motion Instance <-> NC-Task 1 SAF/Axes/Axis 3
//     PlcTask Inputs/Main.M3.Axis.NcToPlc <-> Outputs/ToPlc
//     PlcTask Outputs/Main.M3.Axis.PlcToNc <-> Inputs/FromPlc
//   lfe_motion Instance <-> NC-Task 1 SAF/Axes/Axis 30 IM4L0-XTES-CLF
//     PlcTask Inputs/Main.M30.Axis.NcToPlc <-> Outputs/ToPlc
//     PlcTask Outputs/Main.M30.Axis.PlcToNc <-> Inputs/FromPlc
//   lfe_motion Instance <-> NC-Task 1 SAF/Axes/Axis 33
//     PlcTask Inputs/Main.M33.Axis.NcToPlc <-> Outputs/ToPlc
//     PlcTask Outputs/Main.M33.Axis.PlcToNc <-> Inputs/FromPlc
//   lfe_motion Instance <-> NC-Task 1 SAF/Axes/Axis 34
//     PlcTask Inputs/Main.M34.Axis.NcToPlc <-> Outputs/ToPlc
//     PlcTask Outputs/Main.M34.Axis.PlcToNc <-> Inputs/FromPlc
//   lfe_motion Instance <-> NC-Task 1 SAF/Axes/Axis 35
//     PlcTask Inputs/Main.M35.Axis.NcToPlc <-> Outputs/ToPlc
//     PlcTask Outputs/Main.M35.Axis.PlcToNc <-> Inputs/FromPlc
//   lfe_motion Instance <-> NC-Task 1 SAF/Axes/Axis 36
//     PlcTask Inputs/Main.M36.Axis.NcToPlc <-> Outputs/ToPlc
//     PlcTask Outputs/Main.M36.Axis.PlcToNc <-> Inputs/FromPlc
//   lfe_motion Instance <-> NC-Task 1 SAF/Axes/Axis 37
//     PlcTask Inputs/Main.M37.Axis.NcToPlc <-> Outputs/ToPlc
//     PlcTask Outputs/Main.M37.Axis.PlcToNc <-> Inputs/FromPlc
//   lfe_motion Instance <-> NC-Task 1 SAF/Axes/Axis 38
//     PlcTask Inputs/Main.M38.Axis.NcToPlc <-> Outputs/ToPlc
//     PlcTask Outputs/Main.M38.Axis.PlcToNc <-> Inputs/FromPlc
//   lfe_motion Instance <-> NC-Task 1 SAF/Axes/Axis 39
//     PlcTask Inputs/Main.M39.Axis.NcToPlc <-> Outputs/ToPlc
//     PlcTask Outputs/Main.M39.Axis.PlcToNc <-> Inputs/FromPlc
//   lfe_motion Instance <-> NC-Task 1 SAF/Axes/Axis 4
//     PlcTask Inputs/Main.M4.Axis.NcToPlc <-> Outputs/ToPlc
//     PlcTask Outputs/Main.M4.Axis.PlcToNc <-> Inputs/FromPlc
//   lfe_motion Instance <-> NC-Task 1 SAF/Axes/Axis 40
//     PlcTask Inputs/Main.M40.Axis.NcToPlc <-> Outputs/ToPlc
//     PlcTask Outputs/Main.M40.Axis.PlcToNc <-> Inputs/FromPlc
//   lfe_motion Instance <-> NC-Task 1 SAF/Axes/Axis 5
//     PlcTask Inputs/Main.M5.Axis.NcToPlc <-> Outputs/ToPlc
//     PlcTask Outputs/Main.M5.Axis.PlcToNc <-> Inputs/FromPlc
//   lfe_motion Instance <-> NC-Task 1 SAF/Axes/Axis 6
//     PlcTask Inputs/Main.M6.Axis.NcToPlc <-> Outputs/ToPlc
//     PlcTask Outputs/Main.M6.Axis.PlcToNc <-> Inputs/FromPlc
//   lfe_motion Instance <-> NC-Task 1 SAF/Axes/Axis 7
//     PlcTask Inputs/Main.M7.Axis.NcToPlc <-> Outputs/ToPlc
//     PlcTask Outputs/Main.M7.Axis.PlcToNc <-> Inputs/FromPlc
//   lfe_motion Instance <-> NC-Task 1 SAF/Axes/Axis 8
